(* IEC 61131-3 sources: daoli-st-library/DL_Base (part 5) *)

(* ---- FC_DL_FirstSetBit.st ---- *)
(*==============================================================================
 * 组件名称 (Component)  : FC_DL_FirstSetBit
 * 溯源说明 (Provenance): 道莅 clean-room 防御性实现（IEC 61131-3 纯净实现，闭源文档仅借语义，零代码行）
 * 所属子库 (Sublibrary) : DL_Base / BitString
 * 当前版本 (Version)    : 1.0.0
 * 兼容性   (Platform)   : CODESYS 3.5 / TwinCAT 3 / 汇川 InoProShop / 施耐德
 *                         Machine Expert；纯 IEC 61131-3（第 3 版），仅用
 *                         Standard.library 的 SHR / AND
 * 组件分类 (Category)   : 函数（FUNCTION）· 纯函数 · 位串搜索
 * 功能一句话 (Summary)  : 在 8/16/32/64 位有效位宽内定位**首个置位位**，支持
 *                         低位优先与高位优先两种扫描方向，返回 0 基位号。
 *
 * 本件存在的意义 (Why this unit exists)
 *   位串族已有读写（BitGet/BitSet）、统计（BitCount）、提取（BitFieldExtract）、
 *   批量（BitArray*）、旋转与掩码比较，唯独**搜索**缺位。现场「状态字 →
 *   首个故障位号」「IO 字 → 首个空位」每次都要手写一遍循环，各处写法不一，
 *   64 位宽还有 SHL(x,64) 这类未定义行为的踩坑面。本件把搜索收成一个件。
 *
 * 边界安全 (Boundary)
 *   ① uWidth 不在 {8,16,32,64} → 钳到最近的合法值并置信息 0463（钳位后可继续
 *      工作，属正常防御）；uWidth = 0 → 故障 03B1、bFound = FALSE、bValid = FALSE
 *      （零位宽没有仲裁对象，属非法参数，不是正常结论）；
 *   ② 宽 64 用**常量掩码** DL_MASK64，全程不出现 SHL/SHR 的移位量等于位宽的
 *      写法（R10/R48 两次实证该行为未定义）；移位量恒满足 0 ≤ 移位量 ≤ 63；
 *   ③ 屏蔽后全零 → bFound = FALSE、bValid = TRUE + 信息 0462：「没有置位位」
 *      是合法结论，不是错误；
 *   ④ 高位优先模式下被屏蔽位绝不参与仲裁——先屏蔽、后扫描，顺序不可反；
 *   ⑤ 两个方向都用 WHILE + 守卫计数器（上限 = 有效位宽），超限即退出，
 *      结构性防死锁；高位优先用「步数递增、位号递减」的写法，规避 UINT 下溢。
 * 遗留假设 (Assumption)
 *   LWORD 型 VAR_INPUT 在汇川 InoProShop 的可用性属 P0 编译验证项
 *   （R22 风险表已挂账），本件不降级为 DWORD 双拼，以保持位宽语义完整。
 *
 * 错误码    : 16#0001_0462 屏蔽后全零，无置位位（bFound = FALSE）——信息级，正常结论非错误
 *             16#0001_0463 有效位宽不在 8/16/32/64，已钳位到最近合法值——信息级，正常防御
 *             16#0001_03B1 有效位宽为 0，无法仲裁——故障级，bFound = FALSE 且 bValid = FALSE
 *             16#0001_03B2 预留禁用（故障级，不得挪用）
 *             16#0001_03B3 预留禁用（故障级，不得挪用）
 * 码位总账  : 16#0001_0462 用 / 16#0001_0463 用 ｜ 16#0001_03B1 用 / 16#0001_03B2 预留 / 16#0001_03B3 预留
 * 状态机    : N/A —— 纯函数无顺序状态机
 * 采样约定  : 纯组合函数，无定时器、无内部驻留状态
 * 依赖说明  : 无 DL_ 内部依赖；仅 Standard.library 的 SHR / AND
 * 验收向量  : V1 16#00A0/宽8/低位优先 → uBitIndex=5，bFound=TRUE，TRUE
 *             V2 16#00A0/宽8/高位优先 → uBitIndex=7，bFound=TRUE，TRUE
 *             V3 16#0100/宽8/低位优先 → 屏蔽后全零，bFound=FALSE，bValid=TRUE，eErr=0462，FALSE
 *             V4 16#0100/宽16/低位优先 → uBitIndex=8，bFound=TRUE（掩码边界主向量）
 *             V5 宽 0 → FALSE，eErr=03B1，bValid=FALSE，bError=TRUE
 *             V6 宽 12 → 钳到 16 且 eErr=0463，仍按 16 位仲裁
 *             V7 16#8000_0000_0000_0000/宽64/高位优先 → uBitIndex=63（禁 SHL 64 主向量）
 * 红线自检  : 全局变量声明零使用 / 外部变量访问零使用 / 物理地址零使用 ｜ 纯 IEC 61131-3 ｜ 无除法
 *             无浮点 ｜ 移位量恒小于位宽 ｜ 循环双守卫 ｜ 全变量双语同行注释
 *             状态机 N/A ｜ 无定时器实例 ｜ 掩码与位宽全部常量化
 * 修订历史  : 2026-11-16  v1.0.0  首版入库（R22 · 批 1 · 位串族第四轴）
 *============================================================================*)

FUNCTION FC_DL_FirstSetBit : BOOL
VAR_INPUT
    uValue      : LWORD;                       // 待搜索位串，全域有效 / bit string to search, the whole word is readable
    uWidth      : UINT := 64;                  // 有效位宽 [位]，8/16/32/64 / effective width in bits, 8/16/32/64
    bHighFirst  : BOOL := FALSE;               // TRUE 高位优先 / FALSE 低位优先 / TRUE scans from the top, FALSE from the bottom
END_VAR
VAR_OUTPUT
    uBitIndex   : UINT;                        // 首个置位位号，0 基 [位号] / first set bit index, 0-based
    bFound      : BOOL;                        // 是否找到置位位 / whether a set bit was found
    eErr        : UDINT;                       // 错误码，0 表示无错 / error code, 0 means no error
    bError      : BOOL;                        // 故障级标志，仅故障级错误置位 / fault-class flag, set only on fault-level codes
    bValid      : BOOL;                        // 结论可用标志（全零结论亦为可用） / conclusion usable flag, TRUE for an all-zero conclusion too
END_VAR
VAR
    uWUse       : UINT;                        // 生效有效位宽 [位]，已钳位 / effective width after clamping
    uI          : UINT;                        // 当前候选位号 [位号] / candidate bit index
    uSteps      : UINT;                        // 高位优先的步数计数 [步] / step counter for the downward scan
    uGuard      : UINT;                        // 循环守卫计数器 [次] / loop guard counter
    xMask       : LWORD;                       // 有效位宽掩码 [位串] / mask of the effective width
    xMasked     : LWORD;                       // 屏蔽后的位串 [位串] / bit string after masking
END_VAR
VAR CONSTANT
    DL_W8       : UINT := 8;                   // 合法位宽之一 [位] / one of the legal widths
    DL_W16      : UINT := 16;                  // 合法位宽之一 [位] / one of the legal widths
    DL_W32      : UINT := 32;                  // 合法位宽之一 [位] / one of the legal widths
    DL_W64      : UINT := 64;                  // 合法位宽之一 [位] / one of the legal widths
    DL_W_ZERO   : UINT := 0;                   // 位宽零值，用于非法判定 [位] / zero width, used by the illegal test
    DL_MASK8    : LWORD := 16#0000_0000_0000_00FF; // 8 位掩码常量 [位串] / 8-bit mask constant
    DL_MASK16   : LWORD := 16#0000_0000_0000_FFFF; // 16 位掩码常量 [位串] / 16-bit mask constant
    DL_MASK32   : LWORD := 16#0000_0000_FFFF_FFFF; // 32 位掩码常量 [位串] / 32-bit mask constant
    DL_MASK64   : LWORD := 16#FFFF_FFFF_FFFF_FFFF; // 64 位全一掩码常量，替代 SHL(x,64) [位串] / 64-bit all-ones mask, replaces SHL(x,64)
    DL_BIT_ONE  : LWORD := 16#0000_0000_0000_0001; // 位取用的与掩码 [位串] / AND mask used to test a single bit
    DL_ZERO_LW  : LWORD := 16#0000_0000_0000_0000; // 位串零值 [位串] / zero bit string
END_VAR

(*------------------------------------------------------------------------------
 * 段 1｜返回值与输出预置（L1/L9）
 *      Preset the return value and every output
 *-----------------------------------------------------------------------------*)
FC_DL_FirstSetBit := FALSE;                     // 返回值预置未找到 / preset to not found
uBitIndex := 0;                                 // 位号预置 0 [位号] / index preset to zero
bFound    := FALSE;                             // 找到标志预置 FALSE / found flag preset to FALSE
eErr      := 16#0000_0000;                      // 错误码预置无错 / error code preset to none
bError    := FALSE;                             // 故障标志预置 FALSE / fault flag preset to FALSE
bValid    := FALSE;                             // 结论可用预置 FALSE / usable flag preset to FALSE
uWUse     := DL_W64;                            // 位宽预置最大合法值 / width preset to the maximum legal value
xMask     := DL_MASK64;                         // 掩码预置全一 / mask preset to all ones
xMasked   := DL_ZERO_LW;                        // 屏蔽结果预置零 / masked value preset to zero
uI        := 0;                                 // 位号游标预置 0 / index cursor preset to zero
uSteps    := 0;                                 // 步数计数预置 0 / step counter preset to zero
uGuard    := 0;                                 // 守卫预置 0 / guard preset to zero

(*------------------------------------------------------------------------------
 * 段 2｜位宽闸门（零宽属故障级；非标准宽度钳到最近合法值）
 *      Width gate: zero is a fault, non-standard widths clamp to the nearest legal value
 *-----------------------------------------------------------------------------*)
IF uWidth = DL_W_ZERO THEN
    eErr   := 16#0001_03B1;                     // 故障级：零位宽无法仲裁 / fault: zero width, nothing to arbitrate
    bError := TRUE;                             // 置故障标志 / raise the fault flag
    bValid := FALSE;                            // 结论不可用 / conclusion unusable
    bFound := FALSE;                            // 未找到 / not found
    RETURN;                                     // 早退路径已统一后处理 / the early exit is fully post-processed
END_IF

IF uWidth <= DL_W8 THEN
    uWUse := DL_W8;                             // 钳到 8 位 / clamped to eight bits
    IF uWidth <> DL_W8 THEN
        eErr := 16#0001_0463;                   // 信息级：位宽已钳位 / informational: width clamped
    END_IF
ELSIF uWidth <= DL_W16 THEN
    uWUse := DL_W16;                            // 钳到 16 位 / clamped to sixteen bits
    IF uWidth <> DL_W16 THEN
        eErr := 16#0001_0463;                   // 信息级：位宽已钳位 / informational: width clamped
    END_IF
ELSIF uWidth <= DL_W32 THEN
    uWUse := DL_W32;                            // 钳到 32 位 / clamped to thirty-two bits
    IF uWidth <> DL_W32 THEN
        eErr := 16#0001_0463;                   // 信息级：位宽已钳位 / informational: width clamped
    END_IF
ELSE
    uWUse := DL_W64;                            // 钳到 64 位（含 > 64 的越界输入） / clamped to sixty-four bits
    IF uWidth <> DL_W64 THEN
        eErr := 16#0001_0463;                   // 信息级：位宽已钳位 / informational: width clamped
    END_IF
END_IF

(*------------------------------------------------------------------------------
 * 段 3｜掩码选择（常量掩码，绝不出现 SHL/SHR 移位量等于位宽的写法）
 *      Mask selection by constants, never a shift amount equal to the width
 *-----------------------------------------------------------------------------*)
IF uWUse = DL_W8 THEN
    xMask := DL_MASK8;                          // 8 位掩码 / eight-bit mask
ELSIF uWUse = DL_W16 THEN
    xMask := DL_MASK16;                         // 16 位掩码 / sixteen-bit mask
ELSIF uWUse = DL_W32 THEN
    xMask := DL_MASK32;                         // 32 位掩码 / thirty-two-bit mask
ELSE
    xMask := DL_MASK64;                         // 64 位全一掩码 / sixty-four-bit all-ones mask
END_IF

(*------------------------------------------------------------------------------
 * 段 4｜先屏蔽后扫描（顺序不可反：被屏蔽位绝不参与仲裁）
 *      Mask before scanning, the order cannot be reversed
 *-----------------------------------------------------------------------------*)
xMasked := uValue AND xMask;                    // 无效高位一律清零 / invalid high bits cleared

IF xMasked = DL_ZERO_LW THEN
    eErr   := 16#0001_0462;                     // 信息级：全零，无置位位 / informational: all zero, no set bit
    bFound := FALSE;                            // 未找到 / not found
    bValid := TRUE;                             // 「没有置位位」是合法结论 / an all-zero conclusion is legal
    FC_DL_FirstSetBit := FALSE;                 // 返回未找到 / return not found
    RETURN;
END_IF

(*------------------------------------------------------------------------------
 * 段 5｜扫描（两方向各一套守卫：低位升扫 / 高位降扫，降扫用步数规避下溢）
 *      Scan in both directions, each with its own guard, the downward scan counts steps
 *-----------------------------------------------------------------------------*)
IF NOT bHighFirst THEN
    WHILE (NOT bFound) AND (uI < uWUse) AND (uGuard <= uWUse) DO
        IF (SHR(xMasked, uI) AND DL_BIT_ONE) <> DL_ZERO_LW THEN
            bFound    := TRUE;                  // 命中置位位 / a set bit was hit
            uBitIndex := uI;                    // 记录 0 基位号 / record the 0-based index
        ELSE
            uI := uI + 1;                       // 未命中则升位 / advance when not hit
        END_IF
        uGuard := uGuard + 1;                   // 守卫累计，上限即位宽 / guard bounded by the width
    END_WHILE
ELSE
    WHILE (NOT bFound) AND (uSteps < uWUse) AND (uGuard <= uWUse) DO
        uI := uWUse - 1 - uSteps;               // 位号 = 位宽 − 1 − 步数，恒不下溢 / index never underflows
        IF (SHR(xMasked, uI) AND DL_BIT_ONE) <> DL_ZERO_LW THEN
            bFound    := TRUE;                  // 命中置位位 / a set bit was hit
            uBitIndex := uI;                    // 记录 0 基位号 / record the 0-based index
        ELSE
            uSteps := uSteps + 1;               // 未命中则降位 / step down when not hit
        END_IF
        uGuard := uGuard + 1;                   // 守卫累计 / guard incremented
    END_WHILE
END_IF

(*------------------------------------------------------------------------------
 * 段 6｜出口（未命中属结构性不可达，复用 0462 兜底，R90 不加码）
 *      Exit: a miss is structurally unreachable, the fallback reuses 0462
 *-----------------------------------------------------------------------------*)
IF NOT bFound THEN
    eErr   := 16#0001_0462;                     // 兜底复用：无置位位 / fallback reuse: no set bit
    bValid := TRUE;                             // 结论仍可用 / the conclusion is still usable
    uBitIndex := 0;                             // 位号归 0 / index back to zero
    FC_DL_FirstSetBit := FALSE;                 // 返回未找到 / return not found
    RETURN;
END_IF

bValid := TRUE;                                 // 结论可用 / conclusion usable
FC_DL_FirstSetBit := TRUE;                      // 返回找到 / return found
END_FUNCTION

(* ---- FC_DL_FlatWallHeatLossCalc.st ---- *)
(*
  Component : FC_DL_FlatWallHeatLossCalc
  Category  : DL_Base
  Function  : 多层平壁复合导热 + 表面对流：q = ΔT / (Σ(ti/λi) + 1/h)
  Complexity: C2
  开源溯源 : DLF 内部原创（R94 族模板派生）；参考语义来源见 SOURCE_HUNTING_MATRIX.md
  规则遵从 : R1-R16
  契约     : 输入 rTiC 内侧温度 [℃]、rToC 外侧环境温度 [℃]、afThickMm 各层厚度定长数组 [mm]
             （ARRAY[0..3]，未用层填零）、afLambdaWmK 各层导热系数定长数组 [W/(m·K)]、
             nLayers 有效层数 [层]、rHWm2K 外表面换热系数 [W/(m2·K)]、rAreaM2 传热面积 [m2]；
             输出 rFluxWm2 热流密度 [W/m2]、rResistM2KW 总热阻 [m2·K/W]、rPowerW 总散热功率 [W]、
             xValid 有效标志、nFaultCode 故障码。
  边界     : 层数须 1~4；每层厚度须 >0、导热系数须 >0（零厚度或零导热视为组态错误判 9803）；
             换热系数须 >1.0E-6；总热阻为分母须 >1.0E-9；面积须 ≥0；
             数组固定 4 元素，访问前逐元素双边界校验（R4）。
  码位     : 9801 输入非有限（故障级）；9802 层数越界（故障级）；9803 层参数或换热系数越域（故障级）。
*)
FUNCTION FC_DL_FlatWallHeatLossCalc : BOOL
VAR_INPUT
    rTiC        : LREAL := 120.0;                    // 内侧温度 [℃] EN: the inner surface temperature
    rToC        : LREAL := 25.0;                     // 外侧环境温度 [℃] EN: the outer ambient temperature
    afThickMm   : ARRAY[0..3] OF LREAL;              // 各层厚度，未用层填零 [mm] EN: the layer thicknesses, unused layers hold zero
    afLambdaWmK : ARRAY[0..3] OF LREAL;              // 各层导热系数 [W/(m·K)] EN: the layer thermal conductivities
    nLayers     : INT := 2;                          // 有效层数 [层] EN: the number of valid layers
    rHWm2K      : LREAL := 10.0;                     // 外表面换热系数 [W/(m2·K)] EN: the outer surface heat transfer coefficient
    rAreaM2     : LREAL := 1.0;                      // 传热面积 [m2] EN: the heat transfer area
END_VAR
VAR_OUTPUT
    rFluxWm2     : LREAL;                            // 热流密度 [W/m2] EN: the heat flux density
    rResistM2KW  : LREAL;                            // 总热阻 [m2·K/W] EN: the total thermal resistance
    rPowerW      : LREAL;                            // 总散热功率 [W] EN: the total heat loss power
    xValid       : BOOL;                             // 输出可信标志 EN: the outputs are valid
    nFaultCode   : INT;                              // 0=无故障 9801=输入非有限 9802=层数越界 9803=层参数越域 EN: zero none, 9801 non finite, 9802 layer count out of range, 9803 layer parameter out of range
END_VAR
VAR
    xFinAll : BOOL;                                  // 标量浮点入参有限 EN: the scalar floating inputs are finite
    xLayerOk: BOOL;                                  // 各层参数合法 EN: every layer parameter is legal
    i       : INT;                                   // 层循环索引 [层] EN: the layer loop index
    nScan   : INT;                                   // 实际扫描层数 [层] EN: the effective layer scan count
    rRes    : LREAL;                                 // 导热热阻累加器 [m2·K/W] EN: the conduction resistance accumulator
    rRtot   : LREAL;                                 // 总热阻 [m2·K/W] EN: the total resistance
    rFlux   : LREAL;                                 // 热流密度中间值 [W/m2] EN: the interim heat flux
END_VAR
VAR CONSTANT
    DL_FWH_Z       : LREAL := 0.0;                   // 浮点零常量 EN: the floating point zero constant
    DL_FWH_K1000   : LREAL := 1000.0;                // 毫米转米系数 EN: the millimetre to metre factor
    DL_FWH_LAY_MAX : INT := 4;                       // 层数上限 [层] EN: the upper bound of the layer count
    DL_FWH_IDX_MAX : INT := 3;                       // 数组上界索引 [层] EN: the array upper bound index
    DL_FWH_MIN     : LREAL := 1.0E-9;                // 总热阻与换热系数的下限 EN: the lower bound of the total resistance and the transfer coefficient
    DL_FWH_C_BAD   : INT := 9801;                    // 输入非有限 EN: a non finite input
    DL_FWH_C_LAY   : INT := 9802;                    // 层数越界 EN: the layer count is out of range
    DL_FWH_C_PARAM : INT := 9803;                    // 层参数或换热系数越域 EN: a layer parameter or the transfer coefficient is out of range
END_VAR

// 段1｜出口预置
FC_DL_FlatWallHeatLossCalc := FALSE;   // 返回值预置假 EN: preset the return value to false
rFluxWm2 := DL_FWH_Z;                  // 热流预置零 [W/m2] EN: preset the flux to zero
rResistM2KW := DL_FWH_Z;               // 总热阻预置零 [m2·K/W] EN: preset the total resistance to zero
rPowerW := DL_FWH_Z;                   // 功率预置零 [W] EN: preset the power to zero
xValid := FALSE;                       // 有效标志预置假 EN: preset the validity flag to false
nFaultCode := 0;                       // 故障码预置零 EN: preset the fault code to zero

// 段2｜非有限闸：标量入参全列
xFinAll := (rTiC = rTiC) AND ((rTiC - rTiC) = DL_FWH_Z)
        AND (rToC = rToC) AND ((rToC - rToC) = DL_FWH_Z)
        AND (rHWm2K = rHWm2K) AND ((rHWm2K - rHWm2K) = DL_FWH_Z)
        AND (rAreaM2 = rAreaM2) AND ((rAreaM2 - rAreaM2) = DL_FWH_Z);   // 四标量输入有限性 EN: the finiteness of the four scalar inputs
IF NOT xFinAll THEN                                                     // 非有限出口 EN: leave early on a non finite input
    nFaultCode := DL_FWH_C_BAD;                                         // 非有限码 EN: the non finite code
    RETURN;                                                             // 早退 EN: return early
END_IF

// 段3｜层数域闸：1~4，越界一律拒绝访问数组
IF (nLayers < 1) OR (nLayers > DL_FWH_LAY_MAX) THEN                     // 层数域闸 EN: the layer count domain gate
    nFaultCode := DL_FWH_C_LAY;                                         // 层数越界码 EN: the layer count code
    RETURN;                                                             // 早退 EN: return early
END_IF

// 段4｜逐层累加导热热阻，逐层过非有限与正值闸
rRes := DL_FWH_Z;                                                        // 热阻累加器清零 [m2·K/W] EN: clear the resistance accumulator
xLayerOk := TRUE;                                                        // 假定各层合法 EN: assume every layer is legal
nScan := nLayers;                                                        // 扫描层数 [层] EN: the scan count
FOR i := 0 TO nScan - 1 DO                                               // 定长数组循环（层数已证 ≤4） EN: the fixed array loop, the count is proven at most four
    IF (i >= 0) AND (i <= DL_FWH_IDX_MAX) THEN                           // 逐元素双边界校验 EN: the per element bound check
        IF (afThickMm[i] = afThickMm[i]) AND ((afThickMm[i] - afThickMm[i]) = DL_FWH_Z)
           AND (afLambdaWmK[i] = afLambdaWmK[i]) AND ((afLambdaWmK[i] - afLambdaWmK[i]) = DL_FWH_Z)
           AND (afThickMm[i] > DL_FWH_Z) AND (afLambdaWmK[i] > DL_FWH_Z) THEN
            rRes := rRes + (afThickMm[i] / DL_FWH_K1000) / afLambdaWmK[i];   // 累加 t/λ，[m2·K/W] EN: accumulate the thickness over the conductivity
        ELSE
            xLayerOk := FALSE;                                                   // 某层非法 EN: some layer is illegal
        END_IF
    END_IF
END_FOR
IF NOT xLayerOk THEN                                                             // 层参数非法 EN: a layer parameter is illegal
    nFaultCode := DL_FWH_C_PARAM;                                                // 层参数越域码 EN: the layer parameter code
    RETURN;                                                                      // 早退 EN: return early
END_IF

// 段5｜加表面对流热阻并求热流：q = ΔT / (ΣR + 1/h)
IF (ABS(rHWm2K) < DL_FWH_MIN) OR (rAreaM2 < DL_FWH_Z) THEN                       // 换热系数与面积闸 EN: the coefficient and area gate
    nFaultCode := DL_FWH_C_PARAM;                                                // 越域码 EN: the out of range code
    RETURN;                                                                      // 早退 EN: return early
END_IF
rRtot := rRes + (1.0 / rHWm2K);                                                   // 总热阻 [m2·K/W] EN: the total resistance
IF ABS(rRtot) < DL_FWH_MIN THEN                                                   // 总热阻分母下限 EN: the total resistance gate
    nFaultCode := DL_FWH_C_PARAM;                                                 // 越域码 EN: the out of range code
    RETURN;                                                                       // 早退 EN: return early
END_IF
rFlux := (rTiC - rToC) / rRtot;                                                    // 热流密度，正负随温差 [W/m2] EN: the flux carrying the temperature difference sign
IF rFlux <> rFlux THEN                                                            // 结果复检 EN: recheck the result
    nFaultCode := DL_FWH_C_PARAM;                                                 // 复检失败码 EN: the recheck failure code
    RETURN;                                                                       // 早退，出口保持零哨兵 EN: return early with the zero sentinels
END_IF

// 段6｜出口
rFluxWm2 := rFlux;                                                                // 热流密度出口 [W/m2] EN: the flux output
rResistM2KW := rRtot;                                                             // 总热阻出口 [m2·K/W] EN: the total resistance output
rPowerW := rFlux * rAreaM2;                                                       // 总散热功率 [W] EN: the total power
xValid := TRUE;                                                                   // 结果可信 EN: the results are valid
FC_DL_FlatWallHeatLossCalc := TRUE;                                               // 返回真 EN: return true
END_FUNCTION

(* ---- FC_DL_GrayToBinary.st ---- *)
(*==============================================================================
 * 组件名称 (Component)  : FC_DL_GrayToBinary
 * 所属子库 (Sublibrary) : DL_Base
 * 当前版本 (Version)    : 1.0.0
 * 兼容性   (Platform)   : CODESYS 3.5 / TwinCAT 3 / 汇川 InoProShop / Machine Expert
 *                         仅用标准 SHL / SHR / XOR / AND，无厂商方言
 * 功能描述 (Function)   : 绝对值编码器格雷码 → 标准二进制无符号整数的纯映射函数。
 *                         支持 1~32 位可变位宽；位宽越界时"钳位并继续计算"，
 *                         以 bValid=FALSE + uErrorId 告警，绝不返回 0——
 *                         返回 0 会让上位机看到"位置突然归零"的假故障。
 *                         位宽 32 时 SHL(1,32) 属未定义行为，掩码必须特判为全 1。
 * 算法     (Algorithm)  : 递推式 B = G XOR (G>>1) XOR (G>>2) … XOR (G>>(w-1))（递推至第 w−1 项），
 *                         迭代上界 31，天然有界，无需防死锁计数器。
 * 开源溯源 (Origin)     : 原创实现。格雷码递推式为公开经典算法，位宽钳位与移位特判
 *                         为本库针对三平台差异所做的工程加固。
 * 依赖     (Depends)    : 无 DL_ 内部依赖；无标准库功能块依赖
 * 职责边界 (Scope)      : 本函数不负责 360° 编码器的 Excess 偏移补偿。
 *                         调用顺序应为：转二进制 → 减 Excess 偏移 → 乘分辨率系数。
 * 红线自检 (Redline)    : R1 ✓ 零全局变量表与外部变量引用 ｜ R2 ✓ 零物理 IO 地址直写
 *                         R3 ✓ 纯 IEC 61131-3 ｜ R4 ✓ 越界钳位 + SHL(1,32) 特判 + 空循环边界
 *                         R5 ✓ 全变量中英双语同行注释 ｜ R6 N/A（无状态机）｜ R7 N/A（无实例调用）
 * 修订历史 (Revision)   :
 *   2026-11-14  v1.0.0  首版入库（Phase 1 冷启动 · Level 0 批次）
 *============================================================================*)
FUNCTION FC_DL_GrayToBinary : UDINT
VAR_INPUT
    uGrayValue : UDINT;            // 格雷码原始值，高位脏数据由掩码剔除 / Raw Gray code, dirty high bits removed by the mask
    uBitWidth  : USINT := 32;      // 有效位宽 1..32，越界按边界钳位 / Valid bit width 1..32, clamped at the boundaries
END_VAR
VAR_OUTPUT
    bValid     : BOOL;             // 位宽合法标志，FALSE 表示参数越界已钳位 / Width valid flag, FALSE means clamped
    uErrorId   : UDINT;            // 故障码，0 = 无故障 / Error code, 0 = no error
END_VAR
VAR
    uBinary    : UDINT;            // 转换结果 / Conversion result
    uMask      : UDINT;            // 位宽掩码，仅保留有效位 / Bit-width mask keeping valid bits only
    uWidth     : USINT;            // 钳位后的有效位宽 / Clamped effective bit width
    nIndex     : USINT;            // 递推索引，值域 1..31 / Recurrence index, range 1..31
END_VAR
VAR CONSTANT
    DL_GRAY_WIDTH_MIN : USINT := 1;    // 最小合法位宽 [bit] / Min legal bit width [bit]
    DL_GRAY_WIDTH_MAX : USINT := 32;   // 最大合法位宽 [bit] / Max legal bit width [bit]
END_VAR

(*------------------------------------------------------------------------------
 * 段 1｜返回值与工作变量预置：任何路径下返回值确定
 *      Initialize return value and working variables for determinism
 *-----------------------------------------------------------------------------*)
FC_DL_GrayToBinary := 16#0000_0000;
bValid             := TRUE;
uErrorId           := 16#0000_0000;
uBinary            := 16#0000_0000;
uMask              := 16#0000_0000;
uWidth             := uBitWidth;

(*------------------------------------------------------------------------------
 * 段 2｜位宽钳位（边界 B1）：钳位后继续计算，不中断、不归零
 *      Width clamping: clamp, then keep computing; never abort, never zero the result
 *      下界 0 与上界 >32 均属参数越界，统一报 16#0001_0001
 *-----------------------------------------------------------------------------*)
IF uBitWidth < DL_GRAY_WIDTH_MIN THEN
    uWidth   := DL_GRAY_WIDTH_MIN;
    bValid   := FALSE;
    uErrorId := 16#0001_0001;
ELSIF uBitWidth > DL_GRAY_WIDTH_MAX THEN
    uWidth   := DL_GRAY_WIDTH_MAX;
    bValid   := FALSE;
    uErrorId := 16#0001_0001;
END_IF

(*------------------------------------------------------------------------------
 * 段 3｜掩码构造（边界 B2）：位宽 32 时特判全 1
 *      Mask construction: special-case to all-ones at width 32
 *      SHL(UDINT#1, 32) 在 IEC 中为未定义行为（CODESYS 得 0、部分平台得 1），
 *      因此必须先判 uWidth >= 32，绝不进入移位语句
 *-----------------------------------------------------------------------------*)
IF uWidth >= DL_GRAY_WIDTH_MAX THEN
    uMask := 16#FFFF_FFFF;
ELSE
    uMask := SHL(UDINT#1, USINT_TO_UDINT(uWidth)) - 16#0000_0001;
END_IF

(*------------------------------------------------------------------------------
 * 段 4｜递推转换（边界 B3/B4）：先掩码再逐级异或右移
 *      Recurrence conversion: mask first, then XOR the shifted word level by level
 *      uWidth = 1 时"FOR 1 TO 0"按 IEC 语义执行零次，天然返回原始值；
 *      必须写成 TO (uWidth - 1)，禁止写成 TO uWidth（会多异或一次 SHR(gray, w)）
 *-----------------------------------------------------------------------------*)
uBinary := uGrayValue AND uMask;

IF uWidth > DL_GRAY_WIDTH_MIN THEN
    FOR nIndex := DL_GRAY_WIDTH_MIN TO (uWidth - DL_GRAY_WIDTH_MIN) DO
        uBinary := uBinary XOR SHR(uGrayValue, USINT_TO_UDINT(nIndex));
    END_FOR;
END_IF

(*------------------------------------------------------------------------------
 * 段 5｜结果掩码（边界 B5）：XOR 链可能带入高位脏数据，末尾再截断一次
 *      Result masking: the XOR chain can pull in dirty high bits, truncate at the end
 *-----------------------------------------------------------------------------*)
uBinary := uBinary AND uMask;

FC_DL_GrayToBinary := uBinary;
END_FUNCTION

(* ---- FC_DL_GrayToByteConv.st ---- *)
// FC_DL_GrayToByteConv v1.0.0
// 开源溯源：来源 brOscatLib / URL https://github.com/iec-oscat-mirror / 许可证 MIT / 借鉴点 BYTE_TO_GRAY 反演语义（移位异或链逐位还原）
(*==============================================================================
 * 功能描述: 格雷码 → 二进制转换（8 位）。采用移位异或链三步反演：
 *           b ^= b>>1; b ^= b>>2; b ^= b>>4，等价于逐位累异或 FOR 循环 8 位的
 *           数学结果，位移量 1/2/4 均小于位宽 8（位移量归一，无越界移位）。
 * 接口契约: 输入 bGray（格雷码字节）；返回二进制字节。
 * 修订历史: 2026-11-23  v1.0.0  R74 首版
 *==============================================================================*)

FUNCTION FC_DL_GrayToByteConv : BYTE
VAR_INPUT
    bGray : BYTE := 16#00;   // 格雷码输入字节 [位域] / Gray-coded input byte
END_VAR
VAR
    bAcc : BYTE;             // 累异或工作字节 [位域] / Accumulating work byte
END_VAR

(* —— 段 0：移位异或链反演（三步覆盖 8 位全部位贡献） —— *)
bAcc := bGray;                              // 工作字节装载格雷码 / Work byte loaded with gray code
bAcc := bAcc XOR SHR(bAcc, 1);              // 第一级：右移 1 位异或（覆盖相邻位） / First stage, shift one
bAcc := bAcc XOR SHR(bAcc, 2);              // 第二级：右移 2 位异或（覆盖隔位） / Second stage, shift two
bAcc := bAcc XOR SHR(bAcc, 4);              // 第三级：右移 4 位异或（覆盖高位） / Third stage, shift four
FC_DL_GrayToByteConv := bAcc;               // 返回二进制结果 / Return binary result

END_FUNCTION

(* ---- FC_DL_HammingDist.st ---- *)
(*
  ==================================================================
  组件名 Component  : FC_DL_HammingDist
  分类   Category   : DL_Base
  版本   Version    : 1.0.0
  功能   Purpose    : 汉明距离：两 LWORD 位串逐位异或后统计 1 的个数（等价
                      popcount），输出 0~64。实现取「逐字节分治」口径：先整字
                      XOR 消除公共位，再按 8 字节循环、每字节 8 位内层计数，
                      双层 FOR 均以常量封顶（8/8），结构性无越界、无死循环；
                      移位量 8*i 最大 56 < 64，满足「移位量先归一」纪律。
  来源   Source     : t2-1-lgf-bitlogic（位逻辑族：借 popcount 分治计数口径，
                      实现零源码复制，全自研）
  互引   Cross-ref  : FC_DL_ReverseBitsLword（同族位序变换原子，上游可先做
                      位序归一再进本件；本件不调用它，仅声明同族关系）
  平台   Platform   : 纯 IEC 61131-3（XOR/SHR/AND/FOR），三平台通用
  依赖   Depends    : 无 DL_ 内部依赖；无标准库定时器
  红线   Redline    : R1 零全局/VAR_EXTERNAL/R2 零 %I/%Q/R3 纯 IEC 标准
                      R4 无除法无浮点（整数域无除零面）/R5 全变量双语同行注释
                      R6 纯函数无状态机（CASE 不适用）/R7 无定时器与沿检测
                      R8 循环界与常量全局部化
  验收   Acceptance : V1 uA=uB → 0 ｜ V2 uA=0,uB=全 1 → 64 ｜
                      V3 uA=16#F0F0..,uB=16#0F0F.. → 64 ｜ V4 单 bit 差 → 1
  变更   Revision   : 2026-11-22  v1.0.0  R66 首版（编码阶段批 1 序 1）
  ==================================================================
*)
FUNCTION FC_DL_HammingDist : UDINT
VAR_INPUT
    uA    : LWORD;  // 位串 A [位串] / bit string A [bits]
    uB    : LWORD;  // 位串 B [位串] / bit string B [bits]
END_VAR
VAR_OUTPUT
    uDist : UDINT;  // 汉明距离，0~64 [位] / Hamming distance, 0 to 64 [bit]
END_VAR
VAR
    uXor  : LWORD;  // 异或工作寄存器 [位串] / xor working register [bits]
    uWork : LWORD;  // 移位后的字节级工作量 [位串] / shifted word for byte extraction [bits]
    uByte : BYTE;   // 当前字节切片 [字节] / current byte slice [byte]
    i     : DINT;   // 外层字节循环变量，0~7 [索引] / outer byte loop index, 0 to 7 [index]
    j     : DINT;   // 内层位循环变量，0~7 [索引] / inner bit loop index, 0 to 7 [index]
END_VAR
VAR CONSTANT
    DHD_BYTE_NUM  : DINT := 8;      // LWORD 字节数，外层循环封顶 [字节] / bytes per LWORD, outer loop bound [byte]
    DHD_BIT_NUM   : DINT := 8;      // 每字节数，内层循环封顶 [位] / bits per byte, inner loop bound [bit]
    DHD_BIT_STEP  : DINT := 8;      // 每字节移位步距，8*i ≤ 56 < 64 [位] / shift step per byte [bit]
    DHD_ZERO      : UDINT := UDINT#0;  // 距离零哨兵 [位] / zero sentinel [bit]
END_VAR

// 段 1｜输出预置 / segment 1, preset the outputs
uDist := DHD_ZERO;              // 距离预置 0 / preset distance to zero
FC_DL_HammingDist := DHD_ZERO;  // 返回值与输出同源（R191 名实双出口）/ the return mirrors the output

// 段 2｜整字异或：公共位归零，仅剩差异位 / segment 2, whole word xor keeps only the differing bits
uXor := uA XOR uB;              // 差异位图 [位串] / the difference bitmap [bits]

// 段 3｜逐字节 popcount：双层常量封顶 FOR / segment 3, per byte popcount with constant bounded loops
FOR i := 0 TO DHD_BYTE_NUM - 1 DO       // 8 字节全覆盖 / all 8 bytes covered
    uWork := SHR(uXor, i * DHD_BIT_STEP);  // 移位量 0/8/../56，恒小于 64，合规归一 / shift amounts stay below 64
    uByte := LWORD_TO_BYTE(uWork);         // 取低 8 位为字节切片 / take the low 8 bits as a byte slice
    FOR j := 0 TO DHD_BIT_NUM - 1 DO       // 字节内 8 位逐位判 / test the 8 bits inside the byte
        IF (uByte AND SHL(BYTE#1, j)) <> BYTE#0 THEN  // 掩码 1 左移 j 位，j ≤ 7 恒在字节域内 / mask one shifted by j stays inside the byte domain
            uDist := uDist + UDINT#1;      // 距离累加，上限 64 由位宽结构性保证 / accumulate, capped at 64 by width
        END_IF
    END_FOR
END_FOR

// 段 4｜返回值落位（与 uDist 同值）/ segment 4, publish the return equal to uDist
FC_DL_HammingDist := uDist;     // 名实双出口 / the named and the returned agree
END_FUNCTION

(* ---- FC_DL_HeatTracePowerCalc.st ---- *)
(*
  Component : FC_DL_HeatTracePowerCalc
  Category  : DL_Base
  Function  : 电伴热功率 = 单位热损 × 安全系数，给出每米功率、总功率与工作电流
  Complexity: C2
  开源溯源 : DLF 内部原创（R94 族模板派生）；参考语义来源见 SOURCE_HUNTING_MATRIX.md
  规则遵从 : R1-R16
  契约     : 输入 rLossWm 单位管长设计热损 [W/m]、rSafetyFactor 安全系数 [-]、
             rLengthM 伴热管长 [m]、rVoltageV 供电电压 [V]、rFactorMax 安全系数上限 [-]；
             输出 rPowerWm 每米伴热功率 [W/m]、rPowerTotalW 总伴热功率 [W]、
             rCurrentA 工作电流 [A]、xFactorHigh 安全系数越域（信息级，按上限取值）、
             xValid 有效标志、nFaultCode 故障码。
  边界     : 热损须 ≥0、管长须 ≥0、安全系数须 ≥1 且不超过上限（越域按上限取值并置信息级标志）；
             电压为分母须 >1.0E-6 [V]，否则电流输出 0（不判故障，允许未接线组态）；
             功率上限反算：1.0E4 [W/m] × 1.0E4 [m] ≤ 1.0E8 [W]，远小于 LREAL 上限，可表。
  码位     : 9801 输入非有限（故障级）；9802 热损、管长或安全系数越域（故障级）。
*)
FUNCTION FC_DL_HeatTracePowerCalc : BOOL
VAR_INPUT
    rLossWm      : LREAL := 40.0;    // 单位管长设计热损 [W/m] EN: the design heat loss per metre of pipe
    rSafetyFactor: LREAL := 1.25;    // 安全系数 [-] EN: the safety factor
    rLengthM     : LREAL := 50.0;    // 伴热管长 [m] EN: the traced pipe length
    rVoltageV    : LREAL := 220.0;   // 供电电压 [V] EN: the supply voltage
    rFactorMax   : LREAL := 2.0;     // 安全系数上限 [-] EN: the upper bound of the safety factor
END_VAR
VAR_OUTPUT
    rPowerWm     : LREAL;            // 每米伴热功率 [W/m] EN: the heat tracing power per metre
    rPowerTotalW : LREAL;            // 总伴热功率 [W] EN: the total heat tracing power
    rCurrentA    : LREAL;            // 工作电流 [A] EN: the operating current
    xFactorHigh  : BOOL;             // 安全系数越域（信息级） EN: the safety factor is out of range, information class only
    xValid       : BOOL;             // 输出可信标志 EN: the outputs are valid
    nFaultCode   : INT;              // 0=无故障 9801=输入非有限 9802=热损或管长或系数越域 EN: zero none, 9801 non finite, 9802 loss, length or factor out of range
END_VAR
VAR
    xFinAll : BOOL;                  // 五输入同时有限 EN: all five inputs are finite
    rFacUse : LREAL;                 // 实际使用的安全系数 [-] EN: the safety factor in use
    rPwm    : LREAL;                 // 每米功率中间值 [W/m] EN: the interim power per metre
    rTotal  : LREAL;                 // 总功率中间值 [W] EN: the interim total power
    rCur    : LREAL;                 // 电流中间值 [A] EN: the interim current
END_VAR
VAR CONSTANT
    DL_HTP_Z      : LREAL := 0.0;    // 浮点零常量 EN: the floating point zero constant
    DL_HTP_ONE    : LREAL := 1.0;    // 浮点壹常量 EN: the floating point one constant
    DL_HTP_MIN    : LREAL := 1.0E-6; // 电压与系数下限 EN: the lower bound of the voltage and the factors
    DL_HTP_C_BAD  : INT := 9801;     // 输入非有限 EN: a non finite input
    DL_HTP_C_RANG : INT := 9802;     // 热损或管长或系数越域 EN: the loss, the length or the factor is out of range
END_VAR

// 段1｜出口预置
FC_DL_HeatTracePowerCalc := FALSE;   // 返回值预置假 EN: preset the return value to false
rPowerWm := DL_HTP_Z;                // 每米功率预置零 [W/m] EN: preset the power per metre to zero
rPowerTotalW := DL_HTP_Z;            // 总功率预置零 [W] EN: preset the total power to zero
rCurrentA := DL_HTP_Z;               // 电流预置零 [A] EN: preset the current to zero
xFactorHigh := FALSE;                // 系数越域标志预置假 EN: preset the factor flag to false
xValid := FALSE;                     // 有效标志预置假 EN: preset the validity flag to false
nFaultCode := 0;                     // 故障码预置零 EN: preset the fault code to zero

// 段2｜非有限闸：五输入全列（上限参与域判，漏则越域判据失效）
xFinAll := (rLossWm = rLossWm) AND ((rLossWm - rLossWm) = DL_HTP_Z)
        AND (rSafetyFactor = rSafetyFactor) AND ((rSafetyFactor - rSafetyFactor) = DL_HTP_Z)
        AND (rLengthM = rLengthM) AND ((rLengthM - rLengthM) = DL_HTP_Z)
        AND (rVoltageV = rVoltageV) AND ((rVoltageV - rVoltageV) = DL_HTP_Z)
        AND (rFactorMax = rFactorMax) AND ((rFactorMax - rFactorMax) = DL_HTP_Z);   // 五输入有限性 EN: the finiteness of all five inputs
IF NOT xFinAll THEN                                                                  // 非有限出口 EN: leave early on a non finite input
    nFaultCode := DL_HTP_C_BAD;                                                      // 非有限码 EN: the non finite code
    RETURN;                                                                          // 早退 EN: return early
END_IF

// 段3｜域闸：热损与管长非负、安全系数 ≥1、上限须 ≥1
IF (rLossWm < DL_HTP_Z) OR (rLengthM < DL_HTP_Z) OR (rSafetyFactor < DL_HTP_ONE)
   OR (rFactorMax < DL_HTP_ONE) THEN
    nFaultCode := DL_HTP_C_RANG;                                                     // 越域码 EN: the out of range code
    RETURN;                                                                          // 早退 EN: return early
END_IF

// 段4｜安全系数域：超上限按上限取值并置信息级标志（不中断功率输出）
IF rSafetyFactor > rFactorMax THEN                                                   // 超上限判据 EN: the upper bound test
    rFacUse := rFactorMax;                                                           // 按上限取值 [-] EN: clamp to the upper bound
    xFactorHigh := TRUE;                                                             // 置信息级标志 EN: raise the information class flag
ELSE
    rFacUse := rSafetyFactor;                                                        // 域内直接使用 [-] EN: use the given factor
END_IF

// 段5｜主体：每米功率 = 热损 × 系数；总功率 = 每米 × 管长；电流按电压折算
rPwm := rLossWm * rFacUse;                                                           // 每米伴热功率 [W/m] EN: the power per metre
rTotal := rPwm * rLengthM;                                                           // 总伴热功率 [W] EN: the total power
IF ABS(rVoltageV) < DL_HTP_MIN THEN                                                  // 电压下限：未接线时电流给零 EN: give zero current when the voltage is unusable
    rCur := DL_HTP_Z;                                                                // 电流给零 [A] EN: give a zero current
ELSE
    rCur := rTotal / rVoltageV;                                                      // 工作电流 [A] EN: the operating current
END_IF

// 段6｜结果复检与出口
IF (rPwm <> rPwm) OR (rTotal <> rTotal) OR (rCur <> rCur) THEN                       // 复检：三路非有限 EN: recheck the three results
    nFaultCode := DL_HTP_C_RANG;                                                     // 复检失败码 EN: the recheck failure code
    RETURN;                                                                          // 早退，出口保持零哨兵 EN: return early with the zero sentinels
END_IF
rPowerWm := rPwm;                                                                    // 每米功率出口 [W/m] EN: the power per metre output
rPowerTotalW := rTotal;                                                              // 总功率出口 [W] EN: the total power output
rCurrentA := rCur;                                                                   // 电流出口 [A] EN: the current output
xValid := TRUE;                                                                      // 结果可信 EN: the results are valid
FC_DL_HeatTracePowerCalc := TRUE;                                                    // 返回真 EN: return true
END_FUNCTION

(* ---- FC_DL_InsulationCriticalRadiusCalc.st ---- *)
(*
  Component : FC_DL_InsulationCriticalRadiusCalc
  Category  : DL_Base
  Function  : 临界保温半径 rc = λ/h，并判定当前外径下加保温是否真的减少散热
  Complexity: C2
  开源溯源 : DLF 内部原创（R94 族模板派生）；参考语义来源见 SOURCE_HUNTING_MATRIX.md
  规则遵从 : R1-R16
  契约     : 输入 rLambdaWmK 保温材料导热系数 [W/(m·K)]、rHWm2K 表面换热系数 [W/(m2·K)]、
             rOuterRadiusMm 当前保温外半径 [mm]；
             输出 rCritRadiusMm 临界半径 [mm]、xEffective 加保温有效（外半径 ≥ 临界半径）、
             xValid 有效标志、nFaultCode 故障码。
  边界     : 换热系数为分母须 >1.0E-6 [W/(m2·K)]；导热系数须 >0；外半径须 ≥0；
             临界半径判据针对小管径场景：外半径小于临界半径时，增加保温反而使散热增大，
             此时 xEffective=FALSE（信息级，不置故障）。
  码位     : 9801 输入非有限（故障级）；9802 换热系数或导热系数越域（故障级）。
*)
FUNCTION FC_DL_InsulationCriticalRadiusCalc : BOOL
VAR_INPUT
    rLambdaWmK    : LREAL := 0.045;   // 保温材料导热系数 [W/(m·K)] EN: the thermal conductivity of the insulation
    rHWm2K        : LREAL := 10.0;    // 表面换热系数 [W/(m2·K)] EN: the surface heat transfer coefficient
    rOuterRadiusMm: LREAL := 80.0;    // 当前保温外半径 [mm] EN: the current insulation outer radius
END_VAR
VAR_OUTPUT
    rCritRadiusMm : LREAL;            // 临界保温半径 [mm] EN: the critical insulation radius
    xEffective    : BOOL;             // 加保温对散热有效 EN: the insulation reduces the heat loss
    xValid        : BOOL;             // 输出可信标志 EN: the outputs are valid
    nFaultCode    : INT;              // 0=无故障 9801=输入非有限 9802=换热或导热系数越域 EN: zero none, 9801 non finite, 9802 transfer coefficient or conductivity out of range
END_VAR
VAR
    xFinAll : BOOL;                   // 三输入同时有限 EN: all three inputs are finite
    rDen    : LREAL;                  // 分母（换热系数） [W/(m2·K)] EN: the divisor, the heat transfer coefficient
    rCrit   : LREAL;                  // 临界半径中间值 [mm] EN: the interim critical radius
END_VAR
VAR CONSTANT
    DL_ICR_Z     : LREAL := 0.0;      // 浮点零常量 EN: the floating point zero constant
    DL_ICR_K1000 : LREAL := 1000.0;   // 米转毫米系数 EN: the metre to millimetre factor
    DL_ICR_MIN   : LREAL := 1.0E-6;   // 换热系数下限 EN: the lower bound of the heat transfer coefficient
    DL_ICR_C_BAD : INT := 9801;       // 输入非有限 EN: a non finite input
    DL_ICR_C_RANG: INT := 9802;       // 换热或导热系数越域 EN: the transfer coefficient or the conductivity is out of range
END_VAR

// 段1｜出口预置
FC_DL_InsulationCriticalRadiusCalc := FALSE;   // 返回值预置假 EN: preset the return value to false
rCritRadiusMm := DL_ICR_Z;                     // 临界半径预置零 [mm] EN: preset the critical radius to zero
xEffective := FALSE;                           // 有效保温标志预置假 EN: preset the effective flag to false
xValid := FALSE;                               // 有效标志预置假 EN: preset the validity flag to false
nFaultCode := 0;                               // 故障码预置零 EN: preset the fault code to zero

// 段2｜非有限闸：三输入全列
xFinAll := (rLambdaWmK = rLambdaWmK) AND ((rLambdaWmK - rLambdaWmK) = DL_ICR_Z)
        AND (rHWm2K = rHWm2K) AND ((rHWm2K - rHWm2K) = DL_ICR_Z)
        AND (rOuterRadiusMm = rOuterRadiusMm) AND ((rOuterRadiusMm - rOuterRadiusMm) = DL_ICR_Z);   // 三输入有限性 EN: the finiteness of all three inputs
IF NOT xFinAll THEN                                                                                  // 非有限出口 EN: leave early on a non finite input
    nFaultCode := DL_ICR_C_BAD;                                                                      // 非有限码 EN: the non finite code
    RETURN;                                                                                          // 早退 EN: return early
END_IF

// 段3｜域闸：换热系数过分母下限、导热系数为正、外半径非负
rDen := rHWm2K;                                                                                       // 取分母 [W/(m2·K)] EN: take the divisor
IF (ABS(rDen) < DL_ICR_MIN) OR (rLambdaWmK <= DL_ICR_Z) OR (rOuterRadiusMm < DL_ICR_Z) THEN            // 域闸 EN: the domain gate
    nFaultCode := DL_ICR_C_RANG;                                                                      // 越域码 EN: the out of range code
    RETURN;                                                                                            // 早退 EN: return early
END_IF

// 段4｜主体：rc = λ/h（单位 m），折毫米输出
rCrit := (rLambdaWmK / rDen) * DL_ICR_K1000;                                                           // 临界半径 [mm] EN: the critical radius in millimetres
IF (rCrit <> rCrit) OR (rCrit < DL_ICR_Z) THEN                                                         // 结果复检 EN: recheck the result
    nFaultCode := DL_ICR_C_RANG;                                                                       // 复检失败码 EN: the recheck failure code
    RETURN;                                                                                            // 早退，出口保持零哨兵 EN: return early with the zero sentinels
END_IF

// 段5｜出口：外半径不小于临界半径才判「加保温有效」
rCritRadiusMm := rCrit;                                                                                // 临界半径出口 [mm] EN: the critical radius output
xEffective := rOuterRadiusMm >= rCrit;                                                                 // 有效性判定（信息级） EN: the effectiveness verdict, information class only
xValid := TRUE;                                                                                        // 结果可信 EN: the results are valid
FC_DL_InsulationCriticalRadiusCalc := TRUE;                                                            // 返回真 EN: return true
END_FUNCTION

(* ---- FC_DL_InsulationThicknessCalc.st ---- *)
(*
  Component : FC_DL_InsulationThicknessCalc
  Category  : DL_Base
  Function  : 按单位管长允许热损反求保温层厚度（含表面对流项，不动点迭代 5 次）
  Complexity: C3
  开源溯源 : DLF 内部原创（R94 族模板派生）；参考语义来源见 SOURCE_HUNTING_MATRIX.md
  规则遵从 : R1-R16
  契约     : 输入 rTiC 管内温度 [℃]、rToC 环境温度 [℃]、rLambdaWmK 保温导热系数 [W/(m·K)]、
             rHWm2K 外表面换热系数 [W/(m2·K)]、rInnerDiaMm 保温内径 [mm]、rQallowWm 允许单位热损 [W/m]；
             输出 rThickMm 所需保温厚度 [mm]、rOuterDiaMm 对应保温外径 [mm]、rQcheckWm 代回校验热损 [W/m]、
             xConverged 迭代收敛、xValid 有效标志、nFaultCode 故障码。
  算法     : 串联热阻方程 ln(r2/r1)/(2πλ) + 1/(2π·h·r2) = ΔT/q 无解析解（r2 同时出现在对数与分母），
             故用不动点迭代：r2(k+1) = r1 × exp( 2πλ × (R目标 − 1/(2π·h·r2(k))) )，初值 r2(0)=2·r1，
             固定迭代 5 次（本件迭代次数为常量，不设输入引脚，避免引脚越多验证面越大）。
             收敛判据：代回热损相对误差 ≤1% 判收敛；不收敛仍输出最后一轮值并置 xConverged=FALSE（信息级）。
  边界     : r1 须 >1.0E-4 [mm]、λ 与 h 须 >0、ΔT 须 >0、允许热损须 >0；
             迭代中 r2 若跌破 r1（热阻方程无正解，通常因允许热损大于裸管散热）判 9802。
  码位     : 9801 输入非有限（故障级）；9802 参数越域或无正解（故障级）。
*)
FUNCTION FC_DL_InsulationThicknessCalc : BOOL
VAR_INPUT
    rTiC        : LREAL := 150.0;    // 管内介质温度 [℃] EN: the medium temperature inside the pipe
    rToC        : LREAL := 25.0;     // 环境温度 [℃] EN: the ambient temperature
    rLambdaWmK  : LREAL := 0.045;    // 保温材料导热系数 [W/(m·K)] EN: the thermal conductivity of the insulation
    rHWm2K      : LREAL := 10.0;     // 外表面换热系数 [W/(m2·K)] EN: the outer surface heat transfer coefficient
    rInnerDiaMm : LREAL := 108.0;    // 保温内径（管外径） [mm] EN: the insulation inner diameter, the pipe outer diameter
    rQallowWm   : LREAL := 40.0;     // 允许单位管长热损 [W/m] EN: the allowed heat loss per metre of pipe
END_VAR
VAR_OUTPUT
    rThickMm    : LREAL;             // 所需保温厚度 [mm] EN: the required insulation thickness
    rOuterDiaMm : LREAL;             // 对应保温外径 [mm] EN: the corresponding insulation outer diameter
    rQcheckWm   : LREAL;             // 代回校验的单位热损 [W/m] EN: the heat loss recomputed from the found thickness
    xConverged  : BOOL;              // 迭代收敛（信息级） EN: the iteration converged, information class only
    xValid      : BOOL;              // 输出可信标志 EN: the outputs are valid
    nFaultCode  : INT;               // 0=无故障 9801=输入非有限 9802=参数越域或无正解 EN: zero none, 9801 non finite, 9802 parameters out of range or no positive solution
END_VAR
VAR
    xFinAll : BOOL;                  // 六个浮点入参有限 EN: all six floating inputs are finite
    i       : INT;                   // 迭代计数 [次] EN: the iteration counter
    rR1     : LREAL;                 // 内半径 [m] EN: the inner radius in metres
    rR2     : LREAL;                 // 外半径迭代值 [m] EN: the iterated outer radius
    rRprev  : LREAL;                 // 上一轮外半径 [m] EN: the previous outer radius
    rRtgt   : LREAL;                 // 目标总热阻 [m·K/W] EN: the target total resistance
    rRes    : LREAL;                 // 代回总热阻 [m·K/W] EN: the recomputed total resistance
    rQ      : LREAL;                 // 代回热损 [W/m] EN: the recomputed heat loss
    rErr    : LREAL;                 // 相对误差 [-] EN: the relative error
END_VAR
VAR CONSTANT
    DL_ITC_Z       : LREAL := 0.0;                  // 浮点零常量 EN: the floating point zero constant
    DL_ITC_TWO     : LREAL := 2.0;                  // 直径转半径与初值倍数 EN: the factor used for the radius and the initial guess
    DL_ITC_PI2     : LREAL := 6.2831853071795865;   // 2π（LREAL 精度） [-] EN: twice the circle ratio at LREAL precision
    DL_ITC_K1000   : LREAL := 1000.0;               // 米转毫米系数 EN: the metre to millimetre factor
    DL_ITC_ITER    : INT := 5;                      // 固定迭代次数 [次] EN: the fixed iteration count
    DL_ITC_TOL     : LREAL := 0.01;                 // 收敛相对容差 [-] EN: the convergence tolerance
    DL_ITC_MIN     : LREAL := 1.0E-4;               // 半径下限 [mm] EN: the lower bound of the radius
    DL_ITC_C_BAD   : INT := 9801;                   // 输入非有限 EN: a non finite input
    DL_ITC_C_RANGE : INT := 9802;                   // 参数越域或无正解 EN: parameters out of range or no positive solution
END_VAR

// 段1｜出口预置
FC_DL_InsulationThicknessCalc := FALSE;   // 返回值预置假 EN: preset the return value to false
rThickMm := DL_ITC_Z;                     // 厚度预置零 [mm] EN: preset the thickness to zero
rOuterDiaMm := DL_ITC_Z;                  // 外径预置零 [mm] EN: preset the outer diameter to zero
rQcheckWm := DL_ITC_Z;                    // 校验热损预置零 [W/m] EN: preset the checked loss to zero
xConverged := FALSE;                      // 收敛标志预置假 EN: preset the convergence flag to false
xValid := FALSE;                          // 有效标志预置假 EN: preset the validity flag to false
nFaultCode := 0;                          // 故障码预置零 EN: preset the fault code to zero

// 段2｜非有限闸：六输入全列
xFinAll := (rTiC = rTiC) AND ((rTiC - rTiC) = DL_ITC_Z)
        AND (rToC = rToC) AND ((rToC - rToC) = DL_ITC_Z)
        AND (rLambdaWmK = rLambdaWmK) AND ((rLambdaWmK - rLambdaWmK) = DL_ITC_Z)
        AND (rHWm2K = rHWm2K) AND ((rHWm2K - rHWm2K) = DL_ITC_Z)
        AND (rInnerDiaMm = rInnerDiaMm) AND ((rInnerDiaMm - rInnerDiaMm) = DL_ITC_Z)
        AND (rQallowWm = rQallowWm) AND ((rQallowWm - rQallowWm) = DL_ITC_Z);   // 六输入有限性 EN: the finiteness of all six inputs
IF NOT xFinAll THEN                                                             // 非有限出口 EN: leave early on a non finite input
    nFaultCode := DL_ITC_C_BAD;                                                 // 非有限码 EN: the non finite code
    RETURN;                                                                     // 早退 EN: return early
END_IF

// 段3｜域闸：几何与物性参数正值、温差为正（反向传热无解）
rR1 := (rInnerDiaMm / DL_ITC_TWO) / DL_ITC_K1000;                                // 内半径折米 [m] EN: the inner radius in metres
IF (rInnerDiaMm < DL_ITC_MIN) OR (rLambdaWmK <= DL_ITC_Z) OR (rHWm2K <= DL_ITC_Z)
   OR (rQallowWm <= DL_ITC_Z) OR ((rTiC - rToC) <= DL_ITC_Z) THEN
    nFaultCode := DL_ITC_C_RANGE;                                                // 越域码 EN: the out of range code
    RETURN;                                                                      // 早退 EN: return early
END_IF

// 段4｜目标总热阻与不动点迭代（初值 r2 = 2·r1，固定 5 轮）
rRtgt := (rTiC - rToC) / rQallowWm;                                              // 目标总热阻 [m·K/W] EN: the target total resistance
rR2 := DL_ITC_TWO * rR1;                                                         // 迭代初值 [m] EN: the initial guess
FOR i := 1 TO DL_ITC_ITER DO                                                     // 固定 5 轮，计数器常量化 EN: five fixed rounds
    rRprev := rR2;                                                               // 记上一轮 [m] EN: keep the previous value
    IF (rRprev < DL_ITC_MIN) OR (ABS(rRprev) < DL_ITC_MIN) THEN                  // 迭代值失效保护 EN: guard the iterated value
        rR2 := DL_ITC_TWO * rR1;                                                 // 退回初值 [m] EN: fall back to the initial guess
    ELSE
        rR2 := rR1 * EXP(DL_ITC_PI2 * rLambdaWmK * (rRtgt - (1.0 / (DL_ITC_PI2 * rHWm2K * rRprev))));   // 不动点更新 [m] EN: the fixed point update
    END_IF
    IF rR2 <= rR1 THEN                                                           // 无正解保护：外半径必须大于内半径 EN: the outer radius must exceed the inner one
        nFaultCode := DL_ITC_C_RANGE;                                            // 无正解码 EN: the no positive solution code
        RETURN;                                                                  // 早退 EN: return early
    END_IF
END_FOR

// 段5｜代回校验：q = ΔT / (ln(r2/r1)/(2πλ) + 1/(2π·h·r2))
rRes := LN(rR2 / rR1) / (DL_ITC_PI2 * rLambdaWmK) + (1.0 / (DL_ITC_PI2 * rHWm2K * rR2));   // 代回总热阻 [m·K/W] EN: the recomputed total resistance
IF ABS(rRes) < DL_ITC_TOL THEN                                                             // 热阻下限保护 EN: guard the resistance magnitude
    nFaultCode := DL_ITC_C_RANGE;                                                          // 越域码 EN: the out of range code
    RETURN;                                                                                // 早退 EN: return early
END_IF
rQ := (rTiC - rToC) / rRes;                                                                // 代回热损 [W/m] EN: the recomputed heat loss
rErr := ABS(rQ - rQallowWm) / rQallowWm;                                                    // 相对误差 [-] EN: the relative error
xConverged := rErr <= DL_ITC_TOL;                                                           // 收敛判据（信息级） EN: the convergence verdict, information class only

// 段6｜出口：厚度与热损两出口同源
rThickMm := (rR2 - rR1) * DL_ITC_K1000;                                                     // 所需厚度 [mm] EN: the required thickness
rOuterDiaMm := DL_ITC_TWO * rR2 * DL_ITC_K1000;                                             // 对应外径 [mm] EN: the outer diameter
rQcheckWm := rQ;                                                                            // 校验热损出口 [W/m] EN: the checked loss output
IF rThickMm <= DL_ITC_Z THEN                                                                // 厚度非正判无解 EN: a non positive thickness means no solution
    nFaultCode := DL_ITC_C_RANGE;                                                           // 无正解码 EN: the no solution code
    RETURN;                                                                                 // 早退（返回假） EN: return false
END_IF
xValid := TRUE;                                                                             // 结果可信 EN: the results are valid
FC_DL_InsulationThicknessCalc := TRUE;                                                       // 返回真 EN: return true
END_FUNCTION

(* ---- FC_DL_IntCeilDiv.st ---- *)
(*==============================================================================
 * 组件名称 (Component)  : FC_DL_IntCeilDiv
 * 所属子库 (Sublibrary) : DL_Base
 * 当前版本 (Version)    : 1.0.0
 * 兼容性   (Platform)   : CODESYS 3.5+ / TwinCAT 3 / 汇川 InoProShop / 施耐德 Machine Expert
 *                         仅用标准 / 与 MOD 运算、LINT 中间量，无任何厂商内建函数
 * 功能描述 (Function)   : 整数向上取整除法（向 +∞ 取整，DINT 域）。返回 ceil(nDividend / nDivisor)，
 *                         即满足 nResult × nDivisor >= nDividend 的最小整数（nDivisor > 0 时）。
 *                         用于"件数 = ceil(总长 / 单件长)"、"拍数 = ceil(行程 / 步距)"一类分配
 *                         计算——这类场景必须向上取整，写 (a/b)+1 在整除时会多算一件。
 * 负 数 语 义 (Negative): 本件严格按数学 ceil 定义实现，对负数同样向 +∞ 取整，与截断除法
 *                         （向 0 取整）在异号与同负两种情形下都不同：
 *                           ceil( 7 / 2) =  4  ｜ ceil(-7 / 2) = -3
 *                           ceil( 7 / -2) = -3 ｜ ceil(-7 / -2) =  4
 *                         判据写成"余数与除数同号则商加一"，因此对除数负号同样成立；
 *                         若调用方需要"向 0 取整"或"向 −∞ 取整"，请显式换用本件的兄弟实现，
 *                         不要靠改符号位硬凑（负号外提会改变取整方向）。
 * 已知缺陷对照 (AntiPattern): 禁写 TRUNC(x) + 1 —— ① x 已整除时多算一件；② REAL 域大数精度
 *                         丢失后 TRUNC 结果跳变；③ 负数时 TRUNC 向 0 取整，+1 后方向仍错。
 *                         本件全整数域运算，无 TRUNC、无实数转换，三个缺陷同时规避。
 * 接口     (Interface)  : 入 nDividend 被除数、nDivisor 除数；出 bValid 结果有效、
 *                         bDivZero 除零命中、bOverflow 结果越 DINT 域（已饱和）。
 * 边界     (Boundary)   : ① 除零：不计算，返回 0，bValid=FALSE、bDivZero=TRUE（不抛异常，
 *                         不返回魔数 1 或 −1）；② 溢出：用 LINT 中间量算商，越 DINT 域时
 *                         按符号饱和到 DINT 上下限并置 bOverflow、bValid=FALSE（饱和值可直接
 *                         参与后续比较，但不得当作正确值入库）；③ 无状态：纯组合逻辑，
 *                         同一输入永远同一输出，可任意并发调用（无跨拍驻留）。
 * 依赖     (Depends)    : 无 DL_ 内部依赖；无标准库功能块依赖（仅运算符与类型转换函数）
 * 来源标签 (Source Tag) : T0 防御包装 —— 本件是 **IEC 61131-3 标准语义的道莅防御性实现**：
 *                         向上取整属标准算术语义，防御点在于除零闸、LINT 中间量防溢出、
 *                         余数同号判据（替代 TRUNC+1 缺陷写法）。
 * 码表     (Codes)      : 本件不占用任何全局数字码位。异常出口为 BOOL 三枚
 *                         （bValid / bDivZero / bOverflow）；数字码位待主控收口阶段统一派号。
 * 红线自检 (Redline)    : R1 ✓ 零 GVL/VAR_EXTERNAL ｜ R2 ✓ 零 %I/%Q/%M ｜ R3 ✓ 纯 IEC 61131-3
 *                         R4 ✓ 除零闸 + 溢出双侧直比 + 无浮点比较 ｜ R5 ✓ 声明逐行同行双语注释
 *                         R6 N/A（无状态机，无 CASE） ｜ R7 N/A（无实例调用）
 * 修订历史 (Revision)   : 2026-11-19  v1.0.0  R46 首版（批次 1 · 序号 3）
 *==============================================================================*)
FUNCTION FC_DL_IntCeilDiv : DINT
VAR_INPUT
    nDividend : DINT := 0;      // 被除数（可为负） [无量纲] / Dividend, may be negative [dimensionless]
    nDivisor  : DINT := 1;      // 除数（可为负，0 触发除零闸） [无量纲] / Divisor, may be negative, 0 trips the divide gate
END_VAR
VAR_OUTPUT
    bValid    : BOOL;           // 结果有效（未除零且未溢出） [-] / Result valid, no divide-by-zero and no overflow
    bDivZero  : BOOL;           // 除零命中，返回值为 0 的哨兵 [-] / Division by zero hit, 0 returned as sentinel
    bOverflow : BOOL;           // 结果越 DINT 域，返回值已饱和 [-] / Result out of DINT range, saturated
END_VAR
VAR
    n64Dividend : LINT;         // 被除数的 64 位副本（防 DINT 域内中间溢出） [无量纲] / 64-bit copy of the dividend
    n64Divisor  : LINT;         // 除数的 64 位副本（防 DINT 域内中间溢出） [无量纲] / 64-bit copy of the divisor
    n64Quot     : LINT;         // 截断商（向 0 取整），再按余数修正 [无量纲] / Truncated quotient before remainder correction
    n64Rem      : LINT;         // 余数，符号随被除数（IEC MOD 语义） [无量纲] / Remainder, sign follows the dividend per IEC MOD
END_VAR
VAR CONSTANT
    DL_ICD_DINT_MAX : LINT := 2147483647;    // DINT 上限，饱和基准 [无量纲] / DINT upper bound for saturation
    DL_ICD_DINT_MIN : LINT := -2147483648;   // DINT 下限，饱和基准 [无量纲] / DINT lower bound for saturation
END_VAR

(* —— 段 1：返回值与出口初始化（任何路径下返回值确定） —— *)
FC_DL_IntCeilDiv := 0;              // 缺省返回 0（哨兵，不作正确值解读） / Default 0 sentinel, not a valid answer
bValid           := TRUE;           // 先假定有效，闸门命中时改判 / Assume valid, gates may overrule
bDivZero         := FALSE;          // 除零标志清零 / Divide-by-zero flag cleared
bOverflow        := FALSE;          // 溢出标志清零 / Overflow flag cleared

(* —— 段 2：除零闸（除零是小概率但后果为停机，故前置硬闸并非后置判断） —— *)
IF nDivisor = 0 THEN
    bValid   := FALSE;              // 结果无效 / Result invalid
    bDivZero := TRUE;               // 除零命中 / Divide-by-zero hit
    RETURN;                         // 提前返回，返回值为段 1 的 0 哨兵 / Early return with the 0 sentinel
END_IF

(* —— 段 3：64 位域截断除 + 余数同号进位（数学 ceil 判据，替代 TRUNC+1） —— *)
n64Dividend := DINT_TO_LINT(nDividend);      // 升域防中间溢出 / Widen to avoid intermediate overflow
n64Divisor  := DINT_TO_LINT(nDivisor);       // 升域防中间溢出 / Widen to avoid intermediate overflow
n64Quot     := n64Dividend / n64Divisor;     // 截断商（向 0 取整） / Truncated quotient toward zero
n64Rem      := n64Dividend MOD n64Divisor;   // 余数，符号随被除数 / Remainder, sign of dividend
IF (n64Rem <> 0)                                     // 非整除才可能进位 / Carry only when not exactly divisible
   AND (((n64Rem > 0) AND (n64Divisor > 0))           // 同正：向 +∞ 进位 / Both positive: carry up
     OR ((n64Rem < 0) AND (n64Divisor < 0))) THEN     // 同负：向 +∞ 进位 / Both negative: carry up
    n64Quot := n64Quot + 1;                          // 唯一进位点，全件仅此一处 / The only carry site in this unit
END_IF

(* —— 段 4：越界双侧直比（禁 ABS 单侧——ABS(DINT_MIN) 无符号可表性已失） —— *)
IF (n64Quot > DL_ICD_DINT_MAX) OR (n64Quot < DL_ICD_DINT_MIN) THEN
    bOverflow := TRUE;              // 溢出标志 / Overflow flag
    bValid    := FALSE;             // 结果无效 / Result invalid
    IF n64Quot > 0 THEN
        FC_DL_IntCeilDiv := 2147483647;     // 正溢出饱和到 DINT 上限 / Saturate to DINT max
    ELSE
        FC_DL_IntCeilDiv := -2147483648;    // 负溢出饱和到 DINT 下限 / Saturate to DINT min
    END_IF
    RETURN;                         // 饱和值可参与比较，但不得当正确值 / Saturated value must not be treated as correct
END_IF

(* —— 段 5：正常出口（无隐式转换，显式降域） —— *)
FC_DL_IntCeilDiv := LINT_TO_DINT(n64Quot);   // 已知在域内，显式降域 / Known in range, explicit narrowing
bValid           := TRUE;                    // 结果有效 / Result valid

END_FUNCTION

(* ---- FC_DL_IntFloorDiv.st ---- *)
(*==============================================================================
 * 组件名称 (Component)  : FC_DL_IntFloorDiv
 * 所属子库 (Sublibrary) : DL_Base
 * 当前版本 (Version)    : 1.0.0
 * 兼容性   (Platform)   : CODESYS 3.5+ / TwinCAT 3 / 汇川 InoProShop / 施耐德 Machine Expert
 *                         仅依赖 IEC 61131-3 内建整数除法，零厂商私有库
 * 功能描述 (Function)   : 整数向下取整除法（floor 语义，向 −∞ 取整）。
 *                         与 R46 已入册的 FC_DL_IntCeilDiv 成对：本件向 −∞，那件向 +∞，
 *                         正数域两者等价、负数域才分道，故负数向量是唯一有效判别样本。
 *                         实现路径：先取 IEC 内建整数除法的截断商（向 0 取整）与余数，
 *                         再按"余数与除数异号"判据把商减 1 —— 绝不用 TRUNC(x)+1 类写法
 *                         （R28/R153 整数进位点反例），也不做浮点中转（避免 2^31 精度丢失）。
 *                         验收向量（整数域精确，无容差）：
 *                           (+7, +2) = +3 ；(−7, +2) = −4 ；(+7, −2) = −4 ；(−7, −2) = +3
 *                           同余向量：(+8, +2) = +4 ；(−8, +2) = −4 （整除不偏移）
 *                           边界向量：(MIN_INT, +1) = MIN_INT ；（MIN_INT, −1) 溢出钳位
 * 接口     (Interface)  : 入 nNum 被除数、nDen 除数；出 FC 返回值（floor 商）、bInvalid
 *                         拒算标志（nDen=0 当拍）、bOverflow 溢出钳位标志。
 * 边界     (Boundary)   : ① **零除闸**：nDen = 0 → 返回 0 + bInvalid 当拍，不做任何算术；
 *                         ② **溢出闸**：MIN_INT ÷ −1 在补码域不可表（真值 +2147483648），
 *                         钳位返回 MIN_INT + bOverflow（与 FC_DL_IntCeilDiv 同口径，不饱和到 MAX）；
 *                         ③ 中间量 nQ*nDen 不会溢出：|q·d| ≤ |n| 恒成立，仅 MIN_INT/−1 例外已被②拦截；
 *                         ④ 纯函数无记忆量，无锁存、无跨拍状态；⑤ 零全局耦合、零物理地址。
 * 分工声明 (Scope)      : 本件只管"整数域 floor 商"。不接管：浮点取整（用标准库 TRUNC/FLOOR 包装件）、
 *                         向上取整（属 FC_DL_IntCeilDiv）、取模（属 FC_DL_ModLrealSafe 族）。
 * 来源标签 (Source Tag) : T0 防御包装 —— IEC 61131-3 标准语义的道莅防御性实现
 * 码表     (Codes)      : 本件不占用任何全局数字码位（零码位范式 R297）；诊断由 BOOL 出口承担。
 * 红线自检 (Redline)    : R1 ✓ 零 GVL/VAR_EXTERNAL ｜ R2 ✓ 零 %I/%Q/%M ｜ R3 ✓ 纯 IEC 61131-3
 *                         R4 ✓ 零除闸 + 溢出双侧钳位 ｜ R5 ✓ 声明逐行同行双语注释
 *                         R6 ✓ 判别用 IF/RETURN 链无状态机（无 CASE 需求，非状态件）
 *                         R7 ✓ 无定时器/沿实例（纯组合函数）
 * 修订历史 (Revision)   : 2026-11-19  v1.0.0  R47 首版（批次 1 · 序号 1）
 *==============================================================================*)

FUNCTION FC_DL_IntFloorDiv : DINT
VAR_INPUT
    nNum : DINT := 0;                       // 被除数，全 DINT 域 [-] / Dividend, full DINT domain
    nDen : DINT := 1;                       // 除数，零值拒算 [-] / Divisor, zero value rejected
END_VAR
VAR_OUTPUT
    bInvalid  : BOOL := FALSE;              // 拒算标志（nDen=0，当拍有效） [-] / Rejection flag (nDen=0, this scan)
    bOverflow : BOOL := FALSE;              // 溢出钳位标志（MIN_INT/−1） [-] / Overflow clamp flag
END_VAR
VAR
    nQ : DINT := 0;                         // 截断商中间量（向 0 取整） [-] / Truncated quotient (towards zero)
    nR : DINT := 0;                         // 截断余数中间量（与被除数同号） [-] / Truncated remainder, sign of dividend
END_VAR
VAR CONSTANT
    DL_DINT_MIN : DINT := -2147483647 - 1;  // DINT 最小值（避字面量溢出写法） [-] / DINT minimum, literal-overflow safe
    DL_DINT_MAX : DINT := 2147483647;       // DINT 最大值（上溢反算参照） [-] / DINT maximum, upper-bound reference
END_VAR

(* —— 段 1：返回值与两标志预置（R45 四段式第①段） —— *)
FC_DL_IntFloorDiv := 0;                     // 返回值预置安全值 0 / Return value preset to 0
bInvalid  := FALSE;                         // 拒算标志预置 / Rejection flag preset
bOverflow := FALSE;                         // 溢出标志预置 / Overflow flag preset

(* —— 段 2：域闸门早退（零除，不进入任何算术） —— *)
IF nDen = 0 THEN
    bInvalid := TRUE;                       // 零除拒算 / Division by zero rejected
    FC_DL_IntFloorDiv := 0;                 // 拒算返回值 0 / Return 0 on rejection
    RETURN;                                 // 早退，不委托内建除法 / Early return, built-in division not invoked
END_IF

(* —— 段 3：溢出闸（补码域不可表的唯一象限） —— *)
IF (nNum = DL_DINT_MIN) AND (nDen = -1) THEN
    bOverflow := TRUE;                      // 溢出标志 / Overflow flag
    FC_DL_IntFloorDiv := DL_DINT_MIN;       // 钳位返回 MIN_INT（不饱和到 MAX，保持符号侧一致） / Clamp to MIN_INT
    RETURN;                                 // 早退 / Early return
END_IF

(* —— 段 4：委托内建截断除法取商与余数 —— *)
nQ := nNum / nDen;                          // IEC 整数除法截断（向 0） / IEC integer division truncates towards zero
nR := nNum - nQ * nDen;                     // 余数＝被除数−商×除数（与被除数同号） / Remainder, same sign as dividend

(* —— 段 5：向 −∞ 修正（余数与除数异号则商减 1；整除时 nR=0 不偏移） —— *)
IF (nR <> 0) AND ((nR < 0) <> (nDen < 0)) THEN
    nQ := nQ - 1;                           // 向下取整修正 / Floor correction
END_IF

(* —— 段 6：统一出口（结果复检：商域必在 [MIN_INT, MAX] 内，无需再钳） —— *)
FC_DL_IntFloorDiv := nQ;                    // 输出 floor 商 / Output the floor quotient

END_FUNCTION

(* ---- FC_DL_LeapYearChk.st ---- *)
(*
    FC_DL_LeapYearChk —— 闰年判定原子
    ------------------------------------------------------------------
    分类      : DL_Base / Calendar
    前缀      : FC_DL_
    版本      : 1.0.0
    溯源      : IEC 61131-3 标准语义的道莅防御性实现（格里高利历闰年判定，纯整数四级取余）；
                判定律与库内 FB_DL_YearWindowCheck 的闰年判定同源同序（库内复用，
                不另立第四套闰年律）；年份窗口闸、双律/三律切换、错误分级与码位 100% 自有；
                clean-room 重写，未复制任何闭源厂商源码，参考实现仅限 MIT/Apache 许可
    平台      : 纯 IEC 61131-3，CODESYS V3.5+ / TwinCAT 3 / InoProShop 通用
    作者      : 道莅代码库 · PLC编程专家（R20）
    ------------------------------------------------------------------
    功能说明  : 质保期、维护周期、年度检定、闰日补偿都要先回答「这一年二月有没有 29 号」。
                本件把这个判定从 FB_DL_YearWindowCheck 里抽成原子函数，供日期运算族
                与用户代码直接调用，避免每处各写一遍、各错一处。
                核心防御：① 纯整数取余比较，禁浮点、禁除法——(y MOD 4)、（y MOD 100）、
                   （y MOD 400）三个判据全部是非负操作数，不存在负数取余的平台歧义；
                ② 双律/三律由 bFullRule 显式选择，不猜测：
                   两律 (y MOD 4 = 0 且 y MOD 100 <> 0) 是现场最常用口径；
                   三律再加 y MOD 400 = 0，用于跨 2000 年这类整百年的场景。
                   在 1900~2099 窗口内两律与三律只在 2000 年一个点分歧
                   （1900 非闰、2000 是闰），故整百年一律发信息级提示，
                   让调用方知道这一年的结论取决于哪一套律；
                ③ 年份域外直接升故障级，返回 FALSE 且 bValid = FALSE——
                   对域外年份做静默猜测（例如按两律硬算）会把 2100 判成闰年，
                   而 2100 不是闰年，这种错会一路传到质保到期日；
                ④ 结果用 BOOL 返回，bValid 区分「判否」与「判不了」：
                   FALSE 可能是「不是闰年」，也可能是「没判」，两者绝不可混淆。
                职责边界：年度窗口与周期判定归 FB_DL_YearWindowCheck；周次计算归
                FC_DL_WeekOfYearCalc；日期加减归 FC_DL_DateAddDays；本件只管闰年原子判定。
    编译门槛  : 主路径只用 IEC 61131-3 的 MOD 运算符与 UINT 整数比较，
                无内建函数依赖，三平台与任何编译器均无门槛。
    错误码    : 16#0001_0430 整百年（y MOD 100 = 0），两律与三律在此处分歧，结论取决于 bFullRule——信息级，值可用
                16#0001_0431 预留禁用（信息级，不得挪用）
                16#0001_0366 年份超出 1900~2099 窗口——故障级，返回 FALSE，bValid = FALSE
                16#0001_0367 预留（故障级，不得挪用）
                16#0001_0368 预留禁用（故障级，不得挪用）
    码位总账  : 16#0001_0430 用 / 16#0001_0431 预留 ｜ 16#0001_0366 用 / 16#0001_0367 预留 / 16#0001_0368 预留
    状态机    : R6 标注 N/A —— 本组件为纯函数无顺序状态机，无 CASE 可写，非法状态不可能出现
    采样约定  : 本件无定时器、无沿检测、无状态；单拍纯计算，结论与任务周期无关。
                年份是引脚量而非内部锁存，调用方可逐调用传入不同年份。
    修订记录  : 2026-11-16 v1.0.0 首次入库（R20）
*)
FUNCTION FC_DL_LeapYearChk : BOOL
VAR_INPUT
    nYear            : UINT;                  // 待判定年份 [年]，有效域 1900~2099 / year under test [year], valid domain 1900 to 2099
    bFullRule        : BOOL := FALSE;         // FALSE = 两律；TRUE = 四百年律在内的三律 / FALSE uses the two rules, TRUE adds the four hundred year rule
END_VAR
VAR_OUTPUT
    eErr             : UDINT;                 // 错误码，0=正常 / error id, 0=ok
    bError           : BOOL;                  // 故障标志，eErr 为故障级时 TRUE / error flag, TRUE on fault-level eErr
    bValid           : BOOL;                  // 判定是否有效（域外年份为 FALSE，此时返回值不是结论）/ verdict valid, FALSE when the year is out of domain
END_VAR
VAR CONSTANT
    DL_YEAR_MIN      : UINT := 1900;          // 年份窗口下界 [年] / lower bound of the year window [year]
    DL_YEAR_MAX      : UINT := 2099;          // 年份窗口上界 [年] / upper bound of the year window [year]
    DL_YEAR_STEP4    : UINT := 4;             // 四年律取余基数 [年] / modulus of the four year rule [year]
    DL_YEAR_STEP100  : UINT := 100;           // 百年律取余基数 [年] / modulus of the hundred year rule [year]
    DL_YEAR_STEP400  : UINT := 400;           // 四百年律取余基数 [年] / modulus of the four hundred year rule [year]
    DL_UINT_ZERO     : UINT := 0;             // 无符号零常量，避免裸字面量 [年] / unsigned zero constant [year]
END_VAR
VAR
    bLeap            : BOOL;                  // 闰年判定中间结果 / leap year verdict intermediate
    bCentury         : BOOL;                  // 整百年标志，用于提示两律三律分歧 / century flag used by the divergence hint
END_VAR

// 段 1｜返回值与错误状态预置 / segment 1, preset return value and error status
FC_DL_LeapYearChk := FALSE;                   // 故障缺省返回 FALSE（不是闰年）/ fault default returns FALSE, not a leap year
eErr := 0;                                    // 预置无错误 / preset no error
bError := FALSE;                              // 预置无故障 / preset no fault
bValid := FALSE;                              // 预置判定无效，通过闸门后置位 / preset an invalid verdict, set TRUE after the gate
bLeap := FALSE;                               // 判定中间结果预置 / preset the verdict intermediate
bCentury := FALSE;                            // 整百年标志预置 / preset the century flag

// 段 2｜年份窗口闸：域外不猜，直接升故障级 / segment 2, year window gate, never guess
IF (nYear < DL_YEAR_MIN) OR (nYear > DL_YEAR_MAX) THEN
    eErr := 16#0001_0366;                     // 故障级：年份超窗口 / fault level, the year is out of the window
    bError := TRUE;                           // 置故障标志 / raise the error flag
    bValid := FALSE;                          // 判定无效：返回值不是结论 / the verdict is invalid, the return is no conclusion
    FC_DL_LeapYearChk := FALSE;               // 确定缺省值 / deterministic default
    RETURN;                                   // 出口 / exit
END_IF

// 段 3｜两律判定（与库内 FB_DL_YearWindowCheck 同源同序）/ segment 3, the two rule verdict
bLeap := (nYear MOD DL_YEAR_STEP4 = DL_UINT_ZERO)
         AND (nYear MOD DL_YEAR_STEP100 <> DL_UINT_ZERO); // 四年一闰且百年不闰 / divisible by four and not by one hundred

// 段 4｜四百年律（按 bFullRule 显式并入，整百年因此可判为闰）/ segment 4, the four hundred year rule
IF bFullRule THEN
    IF nYear MOD DL_YEAR_STEP400 = DL_UINT_ZERO THEN
        bLeap := TRUE;                        // 四百年一闰，覆盖两律的否定结论 / divisible by four hundred overrides the negative verdict
    END_IF
END_IF

// 段 5｜整百年分歧提示（信息级，不置 bError）/ segment 5, century divergence hint at info level
bCentury := (nYear MOD DL_YEAR_STEP100 = DL_UINT_ZERO);
IF bCentury THEN
    eErr := 16#0001_0430;                     // 信息级：整百年，结论取决于采用两律还是三律 / info level, the verdict depends on the selected rule set
END_IF

// 段 6｜发布结论 / segment 6, publish the verdict
FC_DL_LeapYearChk := bLeap;                   // TRUE = 闰年 [布尔] / TRUE means a leap year [boolean]
bValid := TRUE;                               // 窗口内判定有效 / the verdict inside the window is valid
bError := FALSE;                              // 信息级不置故障（双保险）/ info level never raises a fault, second line of defence
END_FUNCTION

(* ---- FC_DL_LwordToDwords.st ---- *)
(*==============================================================================
 * 名称 : FC_DL_LwordToDwords —— LWORD 拆解为两个 DWORD（本件返回首 DWORD，dwOther 为次字）
 * 分类 / 前缀 / 版本 : DL_Base / FC_DL_ / 1.0.0
 * 溯源 : 开源语义参考（OSCAT/AixOCAT 族，MIT）或 clean-room IEC 实现，未复制源码
 * 平台 : 纯 IEC 61131-3
 * 功能说明 : 将 64 位输入拆为高/低两个 32 位 DWORD。bHiFirst=TRUE 时首字（返回值）
 *            为高 32 位、次字（dwOther）为低 32 位；FALSE 时角色对调。
 *            拆解全程数值语义（移位 + 掩码），不触碰内存字节序。
 *            边界处理：lwIn 全值域合法，高低双字覆盖完整 64 位，无信息丢失。
 * 错误码 : 无故障路径（全值域合法的纯拆解），eErr 恒 0，bValid 恒 TRUE；
 *          16#0001_1A0D 为本件预留码位，当前实现不发出
 * 状态机 : R6 标注 N/A（纯函数无顺序状态，以本节替代 ELSE 兜底）
 * 红线 : R1/R2/R3 ✓ 零全局/零IO/纯IEC ｜ R4 ✓ 移位量=32<64 ｜ R10 ✓ 标准转换 ｜ R11 ✓ 分号收尾 ｜ R15 ✓ 无保留字撞名
 * 修订记录 : 2026-11-23 v1.0.0 首次入库（R76）
 *============================================================================*)
FUNCTION FC_DL_LwordToDwords : DWORD
VAR_INPUT
    lwIn     : LWORD;    // 待拆解的 64 位输入 [位域] / input lword to be split
    bHiFirst : BOOL;     // TRUE=首字取高 32 位 / TRUE when first dword is the high half
END_VAR
VAR_OUTPUT
    dwOther : DWORD;   // 次字（另一半 32 位）/ the other (second) dword
    eErr    : UDINT;   // 故障码，0=正常（本件无故障路径）/ error code, 0=ok (no fault path)
    bError  : BOOL;    // 故障标志，恒 FALSE / error flag, always FALSE
    bValid  : BOOL;    // TRUE=首/次两字均可用，恒 TRUE / TRUE when both dwords are usable
END_VAR
VAR
    _dwHi : DWORD;     // 高 32 位双字 [位域] / high dword
    _dwLo : DWORD;     // 低 32 位双字 [位域] / low dword
END_VAR

eErr   := 16#0000_0000;                      // 故障码清零 / clear error code
bError := FALSE;                             // 故障标志清零 / clear error flag
bValid := TRUE;                              // 本件全值域合法，恒可用 / always valid

_dwHi := LWORD_TO_DWORD(SHR(lwIn, 32));      // 右移 32 位取高双字（移位量 32<64 安全）/ high dword via shift
_dwLo := LWORD_TO_DWORD(lwIn AND 16#0000_0000_FFFF_FFFF);    // 低 32 位掩码后截取 / low dword via mask

IF bHiFirst THEN                             // 首字 = 高 32 位 / first dword is high half
    FC_DL_LwordToDwords := _dwHi;            // 返回首字为高双字 / return high as first
    dwOther := _dwLo;                        // 次字为低双字 / low as other
ELSE                                         // 首字 = 低 32 位 / first dword is low half
    FC_DL_LwordToDwords := _dwLo;            // 返回首字为低双字 / return low as first
    dwOther := _dwHi;                        // 次字为高双字 / high as other
END_IF

END_FUNCTION

(* ---- FC_DL_MapRangeBipolar.st ---- *)
(*
  FC_DL_MapRangeBipolar —— 双极性对称映射，中点偏置
  分类：DL_Base | 复杂度：2 | 轮次：R86
  开源溯源：道莅原创（clean-room 自研，纯 IEC 61131-3 通用算法），无外部代码引用
  许可证：MIT
  职责：把对称双极性输入量程 [fInMin, fInMax]（中点即零点）映射到对称输出量程 [-fOutAmp, +fOutAmp]：
        out = (in - 中点) / (半量程) * 幅值。中点偏置（输入量程中点不为零，如 4..20 mA 对应 12 为中点）自动扣除。
  契约：fIn 输入、fInMin/fInMax 输入端点、fOutAmp 输出幅值（正数，输出范围 = ±幅值）；
        fOut 映射结果；返回 TRUE 表示 fOut 可信。
  边界：① 量程退化校验（容差 DL_MR_EPS）；② fOutAmp 必须 > 0；③ 六个浮点入参逐一非有限闸；
        ④ 除零防护：除以半量程前已过退化闸；零全局、零物理地址、零库件依赖。
*)
FUNCTION FC_DL_MapRangeBipolar : BOOL
VAR_INPUT
    fIn     : LREAL := 0.0;            // 输入值 [输入量程单位] / The input value in the input range unit
    fInMin  : LREAL := 0.0;            // 输入量程下端点 [输入量程单位] / The input range low end
    fInMax  : LREAL := 100.0;          // 输入量程上端点 [输入量程单位] / The input range high end
    fOutAmp : LREAL := 1.0;            // 输出幅值（输出范围 ±幅值） [输出量程单位] / The output amplitude
END_VAR
VAR_OUTPUT
    fOut : LREAL;                      // 映射结果 [输出量程单位] / The mapped value in the output range unit
END_VAR
VAR
    xBad      : BOOL;                  // 参数非法标志 [—] / The parameter invalid flag
    fInClamp  : LREAL;                 // 钳位后的输入 [输入量程单位] / The clamped input value
    fSpanIn   : LREAL;                 // 输入量程跨度（双倍半量程） [输入量程单位] / The input span
    fMid      : LREAL;                 // 输入量程中点 [输入量程单位] / The input range midpoint
    fHalf     : LREAL;                 // 输入半量程 [输入量程单位] / The half span
END_VAR
VAR CONSTANT
    DL_MB_EPS : LREAL := 1.0E-9;       // 浮点比较容差 [-] / The floating point comparison tolerance
    DL_MB_INF : LREAL := 1.0E30;       // 非有限 / 越界判据上限 [-] / The magnitude gate
    DL_MB_Z   : LREAL := 0.0;          // 浮点零常量 [-] / The floating point zero constant
    DL_MB_TWO : LREAL := 2.0;          // 浮点二常量 [-] / The floating point two constant
END_VAR

FC_DL_MapRangeBipolar := FALSE;                           // 返回值预置假 / preset the return false
fOut := DL_MB_Z;                                          // 输出预置零哨兵 / preset the zero sentinel
xBad := FALSE;                                            // 非法标志预置假 / preset the invalid flag false
IF (fIn <> fIn) OR (ABS(fIn) > DL_MB_INF) THEN            // 输入非有限闸 / the input gate
    xBad := TRUE;                                         // 置非法标志 / raise the invalid flag
END_IF
IF (fInMin <> fInMin) OR (ABS(fInMin) > DL_MB_INF) THEN   // 输入下端非有限闸 / the low end gate
    xBad := TRUE;                                         // 置非法标志 / raise the invalid flag
END_IF
IF (fInMax <> fInMax) OR (ABS(fInMax) > DL_MB_INF) THEN   // 输入上端非有限闸 / the high end gate
    xBad := TRUE;                                         // 置非法标志 / raise the invalid flag
END_IF
IF (fOutAmp <> fOutAmp) OR (ABS(fOutAmp) > DL_MB_INF) THEN // 幅值非有限闸 / the amplitude gate
    xBad := TRUE;                                         // 置非法标志 / raise the invalid flag
END_IF
IF fOutAmp <= DL_MB_EPS THEN                              // 幅值非正 / the amplitude is not positive
    xBad := TRUE;                                         // 置非法标志 / raise the invalid flag
END_IF
fSpanIn := fInMax - fInMin;                               // 输入量程跨度 [输入量程单位] / the input span
IF ABS(fSpanIn) < DL_MB_EPS THEN                          // 输入量程退化（除零防护） / the degenerate span
    xBad := TRUE;                                         // 置非法标志 / raise the invalid flag
END_IF
IF NOT xBad THEN                                          // 参数全通过才映射 / map only when all parameters pass
    fMid := (fInMin + fInMax) / DL_MB_TWO;                // 输入量程中点（中点偏置） [输入量程单位] / the midpoint
    fHalf := fSpanIn / DL_MB_TWO;                         // 输入半量程 [输入量程单位] / the half span
    fInClamp := fIn;                                      // 输入接管 [输入量程单位] / take the input value
    IF fInClamp < fInMin THEN                             // 低于下端点 / below the low end
        fInClamp := fInMin;                               // 钳到下端点 [输入量程单位] / clamp to the low end
    END_IF
    IF fInClamp > fInMax THEN                             // 高于上端点 / above the high end
        fInClamp := fInMax;                               // 钳到上端点 [输入量程单位] / clamp to the high end
    END_IF
    fOut := ((fInClamp - fMid) / fHalf) * fOutAmp;        // 对称映射（分母已证非零） [输出量程单位] / the symmetric mapping
    FC_DL_MapRangeBipolar := TRUE;                        // 映射成功 / the mapping succeeded
ELSE
    fOut := DL_MB_Z;                                      // 非法参数输出零哨兵 [输出量程单位] / the sentinel
    FC_DL_MapRangeBipolar := FALSE;                       // 结果不可信 / the result is not valid
END_IF
END_FUNCTION

(* ---- FC_DL_MapRangeClamped.st ---- *)
(*
  FC_DL_MapRangeClamped —— 双端量程映射并对输入钳位
  分类：DL_Base | 复杂度：2 | 轮次：R86
  开源溯源：道莅原创（clean-room 自研，纯 IEC 61131-3 通用算法），无外部代码引用
  许可证：MIT
  职责：把 [fInMin, fInMax] 内的输入线性映射到 [fOutMin, fOutMax]，输入越界时先钳到输入量程端点再映射。
  契约：fIn 输入 [输入量程单位]、fInMin/fInMax 输入量程端点、fOutMin/fOutMax 输出量程端点；
        fOut 映射结果 [输出量程单位]；返回 TRUE 表示 fOut 可信。
  边界：① 量程退化校验 fInMax <> fInMin（容差 DL_MR_EPS），退化时 fOut 给 fOutMin 且返回 FALSE；
        ② 除零防护：除数 fSpanIn 已过退化闸才做除法；③ 六个浮点入参逐一非有限闸；
        ④ 零全局、零物理地址、零库件依赖。
*)
FUNCTION FC_DL_MapRangeClamped : BOOL
VAR_INPUT
    fIn     : LREAL := 0.0;            // 输入值 [输入量程单位] / The input value in the input range unit
    fInMin  : LREAL := 0.0;            // 输入量程下端点 [输入量程单位] / The input range low end
    fInMax  : LREAL := 100.0;          // 输入量程上端点 [输入量程单位] / The input range high end
    fOutMin : LREAL := 0.0;            // 输出量程下端点 [输出量程单位] / The output range low end
    fOutMax : LREAL := 100.0;          // 输出量程上端点 [输出量程单位] / The output range high end
END_VAR
VAR_OUTPUT
    fOut : LREAL;                      // 映射结果 [输出量程单位] / The mapped value in the output range unit
END_VAR
VAR
    xBad     : BOOL;                   // 参数非法标志 [—] / The parameter invalid flag
    fInClamp : LREAL;                  // 钳位后的输入 [输入量程单位] / The clamped input value
    fSpanIn  : LREAL;                  // 输入量程跨度 [输入量程单位] / The input span
    fSpanOut : LREAL;                  // 输出量程跨度 [输出量程单位] / The output span
END_VAR
VAR CONSTANT
    DL_MR_EPS : LREAL := 1.0E-9;       // 浮点比较容差 [-] / The floating point comparison tolerance
    DL_MR_INF : LREAL := 1.0E30;       // 非有限 / 越界判据上限 [-] / The magnitude gate
    DL_MR_Z   : LREAL := 0.0;          // 浮点零常量 [-] / The floating point zero constant
    DL_MR_ONE : LREAL := 1.0;          // 浮点一常量 [-] / The floating point one constant
END_VAR

FC_DL_MapRangeClamped := FALSE;                           // 返回值预置假 / preset the return false
fOut := fOutMin;                                          // 输出预置为输出下端点哨兵 / preset the low end sentinel
xBad := FALSE;                                            // 非法标志预置假 / preset the invalid flag false
IF (fIn <> fIn) OR (ABS(fIn) > DL_MR_INF) THEN            // 输入非有限闸 / the input gate
    xBad := TRUE;                                         // 置非法标志 / raise the invalid flag
END_IF
IF (fInMin <> fInMin) OR (ABS(fInMin) > DL_MR_INF) THEN   // 输入下端非有限闸 / the low end gate
    xBad := TRUE;                                         // 置非法标志 / raise the invalid flag
END_IF
IF (fInMax <> fInMax) OR (ABS(fInMax) > DL_MR_INF) THEN   // 输入上端非有限闸 / the high end gate
    xBad := TRUE;                                         // 置非法标志 / raise the invalid flag
END_IF
IF (fOutMin <> fOutMin) OR (ABS(fOutMin) > DL_MR_INF) THEN // 输出下端非有限闸 / the output low end gate
    xBad := TRUE;                                         // 置非法标志 / raise the invalid flag
END_IF
IF (fOutMax <> fOutMax) OR (ABS(fOutMax) > DL_MR_INF) THEN // 输出上端非有限闸 / the output high end gate
    xBad := TRUE;                                         // 置非法标志 / raise the invalid flag
END_IF
fSpanIn := fInMax - fInMin;                               // 输入量程跨度 [输入量程单位] / the input span
fSpanOut := fOutMax - fOutMin;                            // 输出量程跨度 [输出量程单位] / the output span
IF ABS(fSpanIn) < DL_MR_EPS THEN                          // 输入量程退化（除零防护） / the degenerate input span
    xBad := TRUE;                                         // 置非法标志 / raise the invalid flag
END_IF
IF NOT xBad THEN                                          // 参数全通过才映射 / map only when all parameters pass
    fInClamp := fIn;                                      // 输入接管 [输入量程单位] / take the input value
    IF fSpanIn > DL_MR_Z THEN                             // 正常量程方向 / the normal range direction
        IF fInClamp < fInMin THEN                         // 低于下端点 / below the low end
            fInClamp := fInMin;                           // 钳到下端点 [输入量程单位] / clamp to the low end
        END_IF
        IF fInClamp > fInMax THEN                         // 高于上端点 / above the high end
            fInClamp := fInMax;                           // 钳到上端点 [输入量程单位] / clamp to the high end
        END_IF
    ELSE                                                  // 反向量程（上端小于下端） / the reversed range
        IF fInClamp > fInMin THEN                         // 高于下端点 / above the low end
            fInClamp := fInMin;                           // 钳到下端点 [输入量程单位] / clamp to the low end
        END_IF
        IF fInClamp < fInMax THEN                         // 低于上端点 / below the high end
            fInClamp := fInMax;                           // 钳到上端点 [输入量程单位] / clamp to the high end
        END_IF
    END_IF
    fOut := fOutMin + ((fInClamp - fInMin) / fSpanIn) * fSpanOut; // 线性映射（分母已证非零） [输出量程单位]
    FC_DL_MapRangeClamped := TRUE;                        // 映射成功 / the mapping succeeded
ELSE
    fOut := fOutMin;                                      // 非法参数输出下端点哨兵 [输出量程单位] / the sentinel
    FC_DL_MapRangeClamped := FALSE;                       // 结果不可信 / the result is not valid
END_IF
END_FUNCTION

(* ---- FC_DL_MapRangeDeadband.st ---- *)
(*
  FC_DL_MapRangeDeadband —— 带中心死区的量程映射，死区内输出中点
  分类：DL_Base | 复杂度：2 | 轮次：R86
  开源溯源：道莅原创（clean-room 自研，纯 IEC 61131-3 通用算法），无外部代码引用
  许可证：MIT
  职责：以输入量程中点为中心设置 ±fDbHalf 死区；死区内输出量程中点；
        死区外按「扣除死区后重新归一」的比例映射，保证在死区边界处连续无跳变。
  契约：fIn 输入、fInMin/fInMax 输入端点、fOutMin/fOutMax 输出端点、fDbHalf 死区半宽 [输入量程单位]；
        fOut 映射结果；返回 TRUE 表示可信。
  边界：① 量程与死区退化校验（容差 DL_MD_EPS）；死区半宽必须 >= 0 且 < 输入半量程；
        ② 六个浮点入参逐一非有限闸；③ 除零防护：归一化分母经非退化闸证明 > 0；
        ④ 零全局、零物理地址、零库件依赖。
*)
FUNCTION FC_DL_MapRangeDeadband : BOOL
VAR_INPUT
    fIn     : LREAL := 0.0;            // 输入值 [输入量程单位] / The input value
    fInMin  : LREAL := 0.0;            // 输入量程下端点 [输入量程单位] / The input range low end
    fInMax  : LREAL := 100.0;          // 输入量程上端点 [输入量程单位] / The input range high end
    fOutMin : LREAL := 0.0;            // 输出量程下端点 [输出量程单位] / The output range low end
    fOutMax : LREAL := 100.0;          // 输出量程上端点 [输出量程单位] / The output range high end
    fDbHalf : LREAL := 5.0;            // 死区半宽（以输入中点为心） [输入量程单位] / The dead band half width
END_VAR
VAR_OUTPUT
    fOut  : LREAL;                     // 映射结果 [输出量程单位] / The mapped value
    xInDb : BOOL;                      // 本拍输入落在死区内 [—] / The input is inside the dead band
END_VAR
VAR
    xBad    : BOOL;                    // 参数非法标志 [—] / The parameter invalid flag
    fInMid  : LREAL;                   // 输入量程中点 [输入量程单位] / The input midpoint
    fOutMid : LREAL;                   // 输出量程中点 [输出量程单位] / The output midpoint
    fInHalf : LREAL;                   // 输入半量程 [输入量程单位] / The input half span
    fOutHalf : LREAL;                  // 输出半量程 [输出量程单位] / The output half span
    fRel    : LREAL;                   // 扣除死区后的归一化比例 [归一化] / The normalised ratio beyond the band
    fDev    : LREAL;                   // 输入相对中点的偏移 [输入量程单位] / The deviation from the midpoint
END_VAR
VAR CONSTANT
    DL_MD_EPS  : LREAL := 1.0E-9;      // 浮点比较容差 [-] / The floating point comparison tolerance
    DL_MD_INF  : LREAL := 1.0E30;      // 非有限 / 越界判据上限 [-] / The magnitude gate
    DL_MD_Z    : LREAL := 0.0;         // 浮点零常量 [-] / The floating point zero constant
    DL_MD_TWO  : LREAL := 2.0;         // 浮点二常量 [-] / The floating point two constant
END_VAR

FC_DL_MapRangeDeadband := FALSE;                          // 返回值预置假 / preset the return false
fOut := fOutMin;                                          // 输出预置为输出下端点哨兵 / preset the low end sentinel
xInDb := FALSE;                                           // 死区标志预置假 / preset the dead band flag false
xBad := FALSE;                                            // 非法标志预置假 / preset the invalid flag false
IF (fIn <> fIn) OR (ABS(fIn) > DL_MD_INF) THEN            // 输入非有限闸 / the input gate
    xBad := TRUE;                                         // 置非法标志 / raise the invalid flag
END_IF
IF (fInMin <> fInMin) OR (ABS(fInMin) > DL_MD_INF) THEN   // 输入下端非有限闸 / the input low end gate
    xBad := TRUE;                                         // 置非法标志 / raise the invalid flag
END_IF
IF (fInMax <> fInMax) OR (ABS(fInMax) > DL_MD_INF) THEN   // 输入上端非有限闸 / the input high end gate
    xBad := TRUE;                                         // 置非法标志 / raise the invalid flag
END_IF
IF (fOutMin <> fOutMin) OR (ABS(fOutMin) > DL_MD_INF) THEN // 输出下端非有限闸 / the output low end gate
    xBad := TRUE;                                         // 置非法标志 / raise the invalid flag
END_IF
IF (fOutMax <> fOutMax) OR (ABS(fOutMax) > DL_MD_INF) THEN // 输出上端非有限闸 / the output high end gate
    xBad := TRUE;                                         // 置非法标志 / raise the invalid flag
END_IF
IF (fDbHalf <> fDbHalf) OR (ABS(fDbHalf) > DL_MD_INF) THEN // 死区半宽非有限闸 / the dead band gate
    xBad := TRUE;                                         // 置非法标志 / raise the invalid flag
END_IF
fInHalf := (fInMax - fInMin) / DL_MD_TWO;                 // 输入半量程 [输入量程单位] / the input half span
fOutHalf := (fOutMax - fOutMin) / DL_MD_TWO;              // 输出半量程 [输出量程单位] / the output half span
IF ABS(fInHalf) < DL_MD_EPS THEN                          // 输入量程退化 / the degenerate input span
    xBad := TRUE;                                         // 置非法标志 / raise the invalid flag
END_IF
IF (fDbHalf < DL_MD_Z) OR (ABS(fDbHalf) >= ABS(fInHalf)) THEN // 死区半宽越界 / the dead band is out of range
    xBad := TRUE;                                         // 置非法标志 / raise the invalid flag
END_IF
IF NOT xBad THEN                                          // 参数全通过才映射 / map only when all parameters pass
    fInMid := (fInMin + fInMax) / DL_MD_TWO;              // 输入量程中点 [输入量程单位] / the input midpoint
    fOutMid := (fOutMin + fOutMax) / DL_MD_TWO;           // 输出量程中点 [输出量程单位] / the output midpoint
    fDev := fIn - fInMid;                                 // 输入相对中点偏移 [输入量程单位] / the deviation
    IF ABS(fDev) <= fDbHalf THEN                          // 落在死区内 / inside the dead band
        fOut := fOutMid;                                  // 死区内输出中点 [输出量程单位] / output the midpoint
        xInDb := TRUE;                                    // 置死区标志 [—] / raise the dead band flag
    ELSE
        fRel := (ABS(fDev) - fDbHalf) / (ABS(fInHalf) - ABS(fDbHalf)); // 扣除死区后归一（分母已证 > 0）
        IF fRel > 1.0 THEN                                // 越出量程上界钳位 / clamp beyond the range
            fRel := 1.0;                                  // 钳到一 [归一化] / clamp to one
        END_IF
        IF fDev > DL_MD_Z THEN                            // 正向偏移 / a positive deviation
            fOut := fOutMid + fRel * fOutHalf;            // 正向落位 [输出量程单位] / the positive side
        ELSE
            fOut := fOutMid - fRel * fOutHalf;            // 负向落位 [输出量程单位] / the negative side
        END_IF
    END_IF
    FC_DL_MapRangeDeadband := TRUE;                       // 映射成功 / the mapping succeeded
ELSE
    fOut := fOutMin;                                      // 非法参数输出下端点哨兵 [输出量程单位] / the sentinel
    FC_DL_MapRangeDeadband := FALSE;                      // 结果不可信 / the result is not valid
END_IF
END_FUNCTION

(* ---- FC_DL_MapRangeHystSwitch.st ---- *)
(*
  FC_DL_MapRangeHystSwitch —— 带滞环的二态阈值映射
  分类：DL_Base | 复杂度：2 | 轮次：R86
  开源溯源：道莅原创（clean-room 自研，纯 IEC 61131-3 通用算法），无外部代码引用
  许可证：MIT
  职责：把连续输入映射为两态输出并带滞环：fIn >= fThOn 置态；fIn <= fThOff 复位态；
        fThOff < fIn < fThOn 区间保持上拍态。状态由 VAR_IN_OUT 变量在调用方持有（FC 无内部记忆）。
  契约：fIn 输入、fThOn 置位阈值、fThOff 复位阈值（必须 fThOn > fThOff）、xState 状态输入输出；
        xOut 本拍输出；返回 TRUE 表示可信（参数合法）。
  边界：① 阈值倒置 / 相等校验（容差 DL_MH_EPS）判非法并保持上拍态；② 三个浮点入参非有限闸；
        ③ 滞环区间内显式保持，禁「按当下输入重算」；④ 零全局、零物理地址、零库件依赖。
*)
FUNCTION FC_DL_MapRangeHystSwitch : BOOL
VAR_INPUT
    fIn    : LREAL := 0.0;             // 输入值 [工程单位] / The input value
    fThOn  : LREAL := 80.0;            // 置位阈值（高端） [工程单位] / The set threshold, the high side
    fThOff : LREAL := 20.0;            // 复位阈值（低端） [工程单位] / The reset threshold, the low side
END_VAR
VAR_IN_OUT
    xState : BOOL;                     // 两态状态（调用方持有，跨调用保持） [—] / The two state flag held by the caller
END_VAR
VAR_OUTPUT
    xOut : BOOL;                       // 本拍两态输出 [—] / The two state output
END_VAR
VAR
    xBad : BOOL;                       // 参数非法标志 [—] / The parameter invalid flag
END_VAR
VAR CONSTANT
    DL_MH_EPS : LREAL := 1.0E-9;       // 浮点比较容差 [-] / The floating point comparison tolerance
    DL_MH_INF : LREAL := 1.0E30;       // 非有限 / 越界判据上限 [-] / The magnitude gate
END_VAR

FC_DL_MapRangeHystSwitch := FALSE;                        // 返回值预置假 / preset the return false
xOut := xState;                                           // 输出先保持上拍态 / hold the previous state first
xBad := FALSE;                                            // 非法标志预置假 / preset the invalid flag false
IF (fIn <> fIn) OR (ABS(fIn) > DL_MH_INF) THEN            // 输入非有限闸 / the input gate
    xBad := TRUE;                                         // 置非法标志 / raise the invalid flag
END_IF
IF (fThOn <> fThOn) OR (ABS(fThOn) > DL_MH_INF) THEN      // 置位阈值非有限闸 / the set threshold gate
    xBad := TRUE;                                         // 置非法标志 / raise the invalid flag
END_IF
IF (fThOff <> fThOff) OR (ABS(fThOff) > DL_MH_INF) THEN   // 复位阈值非有限闸 / the reset threshold gate
    xBad := TRUE;                                         // 置非法标志 / raise the invalid flag
END_IF
IF (fThOn - fThOff) < DL_MH_EPS THEN                      // 阈值倒置或相等，滞环宽度非正 / the band is not positive
    xBad := TRUE;                                         // 置非法标志 / raise the invalid flag
END_IF
IF NOT xBad THEN                                          // 参数合法才更新状态 / update only with valid parameters
    IF fIn >= fThOn THEN                                  // 达到置位阈值 / the set threshold is reached
        xState := TRUE;                                   // 置位（滞环高端） [—] / set the state
    ELSIF fIn <= fThOff THEN                              // 达到复位阈值 / the reset threshold is reached
        xState := FALSE;                                  // 复位（滞环低端） [—] / reset the state
    END_IF                                                // 滞环区间内不赋值，xState 自然保持上拍态 / hold inside the band
    xOut := xState;                                       // 状态发布到出口 / publish the state
    FC_DL_MapRangeHystSwitch := TRUE;                     // 参数合法，输出可信 / the parameters are valid
ELSE
    xOut := xState;                                       // 非法参数保持上拍态 [—] / hold the previous state
    FC_DL_MapRangeHystSwitch := FALSE;                    // 结果不可信 / the result is not valid
END_IF
END_FUNCTION
